	            "POS3_0_Signal"."-1002T1 Oriental_Steuerung".E_DDO_Pos := LREAL_TO_REAL("HMI_COM".HMI_Achse_Steuerung.E_Sollwert_Manuell);
	            "POS3_0_Signal"."-1002T1 Oriental_Steuerung".E_Schrittweite := LREAL_TO_REAL("HMI_COM".HMI_Achse_Steuerung.E_Verfahrweg);
	            "POS3_0_Signal"."-1002T1 Oriental_Steuerung".E_DDO_Vel := LREAL_TO_REAL("HMI_COM".HMI_Achse_Steuerung.E_Geschwindigkeit_manuell_in_Prozent);
	            "POS3_0_Signal"."-1002T1 Oriental_Steuerung".E_DDO_Acc := 100.0;
	            "POS3_0_Signal"."-1002T1 Oriental_Steuerung".E_DDO_Dec := 100.0;
	            "POS3_0_Signal"."-1002T1 Oriental_Steuerung".E_DDO_Crnt := 100;
	            
	            "POS3_0_Signal"."-1002T1 Oriental_Steuerung".E_Schrittweite_pos := "HMI_COM".HMI_Achse_Steuerung.E_Tipp_pos;
	            "POS3_0_Signal"."-1002T1 Oriental_Steuerung".E_Schrittweite_neg := "HMI_COM".HMI_Achse_Steuerung.E_Tipp_neg;
	            "POS3_0_Signal"."-1002T1 Oriental_Steuerung".E_Trig_Manuell := "HMI_COM".HMI_Achse_Steuerung.E_Start_manuell;
	            "POS3_0_Signal"."-1002T1 Oriental_Steuerung"."E_FW-JOG" := "HMI_COM".HMI_Achse_Steuerung.E_jog_pos;
	            "POS3_0_Signal"."-1002T1 Oriental_Steuerung"."E_RV-JOG" := "HMI_COM".HMI_Achse_Steuerung.E_jog_neg;
	        //    "HMI_COM".HMI_Achse_Steuerung.E_Start_manuell := false;
	        END_IF;
	       
	            // Initialisieren der Steuerwerte 
	            #R_TRIG_Init_Achse_2_Positionen(CLK := "HMI_SYS"."Aktueller Bildschirm" = #Manuell_Positionen_1_Achse_2);
	        IF #R_TRIG_Init_Achse_2_Positionen.Q THEN
	                "HMI_COM".HMI_Achse_POS_Überschreiben.Wert_Position_Überschreiben[0] := "POS3_0_Signal"."-1002T1 Oriental_Positionen".Soll_Position[0];
	                "HMI_COM".HMI_Achse_POS_Überschreiben.Wert_Speed_Überschreiben[0] := "POS3_0_Signal"."-1002T1 Oriental_Positionen".Geschwindigkeit[0];
	                
	                "HMI_COM".HMI_Achse_POS_Überschreiben.Wert_Position_Überschreiben[1] := "POS3_0_Signal"."-1002T1 Oriental_Positionen".Soll_Position[1];
	                "HMI_COM".HMI_Achse_POS_Überschreiben.Wert_Speed_Überschreiben[1] := "POS3_0_Signal"."-1002T1 Oriental_Positionen".Geschwindigkeit[1];
	                
	                "HMI_COM".HMI_Achse_POS_Überschreiben.Wert_Position_Überschreiben[2] := "POS3_0_Signal"."-1002T1 Oriental_Positionen".Soll_Position[2];
	                "HMI_COM".HMI_Achse_POS_Überschreiben.Wert_Speed_Überschreiben[2] := "POS3_0_Signal"."-1002T1 Oriental_Positionen".Geschwindigkeit[2];
	                
	                "HMI_COM".HMI_Achse_POS_Überschreiben.Wert_Position_Überschreiben[3] := "POS3_0_Signal"."-1002T1 Oriental_Positionen".Soll_Position[3];
	                "HMI_COM".HMI_Achse_POS_Überschreiben.Wert_Speed_Überschreiben[3] := "POS3_0_Signal"."-1002T1 Oriental_Positionen".Geschwindigkeit[3];
	                
	                "HMI_COM".HMI_Achse_POS_Überschreiben.Wert_Position_Überschreiben[4] := "POS3_0_Signal"."-1002T1 Oriental_Positionen".Soll_Position[4];
	                "HMI_COM".HMI_Achse_POS_Überschreiben.Wert_Speed_Überschreiben[4] := "POS3_0_Signal"."-1002T1 Oriental_Positionen".Geschwindigkeit[4];
	                
	                "HMI_COM".HMI_Achse_POS_Überschreiben.Wert_Position_Überschreiben[5] := "POS3_0_Signal"."-1002T1 Oriental_Positionen".Soll_Position[5];
	                "HMI_COM".HMI_Achse_POS_Überschreiben.Wert_Speed_Überschreiben[5] := "POS3_0_Signal"."-1002T1 Oriental_Positionen".Geschwindigkeit[5];
	        END_IF;
	            
	            
	        IF ("HMI_SYS"."Aktueller Bildschirm" = #Manuell_Positionen_1_Achse_2) THEN
	            
	            "HMI_COM".HMI_Achse_Steuerung.A_StatusWord := "POS3_0_Signal"."-1002T1 Oriental_Steuerung".A_StatusWord;
	            "HMI_COM".HMI_Achse_Steuerung.E_Drehachse := false;
	            "HMI_COM".HMI_Achse_Steuerung.A_Istwert := REAL_TO_LREAL("POS3_0_Signal"."-1002T1 Oriental_Steuerung".A_FBposition);
	            "HMI_COM".HMI_Achse_Steuerung.A_Softw_ES_min := "POS3_0_Signal"."-1002T1 Oriental_Positionen".A_Softw_ES_min_mm;
	            "HMI_COM".HMI_Achse_Steuerung.A_Softw_ES_max := "POS3_0_Signal"."-1002T1 Oriental_Positionen".A_Softw_ES_max_mm;
	            
	            
	            "HMI_COM".HMI_Achse_Position.Soll_Wert_in_mm_Position[0] := "POS3_0_Signal"."-1002T1 Oriental_Positionen".Soll_Position[0];
	            "HMI_COM".HMI_Achse_Position.Soll_Wert_in_mm_Position[1] := "POS3_0_Signal"."-1002T1 Oriental_Positionen".Soll_Position[1];
	            "HMI_COM".HMI_Achse_Position.Soll_Wert_in_mm_Position[2] := "POS3_0_Signal"."-1002T1 Oriental_Positionen".Soll_Position[2];
	            "HMI_COM".HMI_Achse_Position.Soll_Wert_in_mm_Position[3] := "POS3_0_Signal"."-1002T1 Oriental_Positionen".Soll_Position[3];
	            "HMI_COM".HMI_Achse_Position.Soll_Wert_in_mm_Position[4] := "POS3_0_Signal"."-1002T1 Oriental_Positionen".Soll_Position[4];
	            "HMI_COM".HMI_Achse_Position.Soll_Wert_in_mm_Position[5] := "POS3_0_Signal"."-1002T1 Oriental_Positionen".Soll_Position[5];
	            
	            "HMI_COM".HMI_Achse_Position.POS_OK_Position[0] := "POS3_0_Signal"."-1002T1 Oriental_Positionen".POS_OK_Position[0];
	            "HMI_COM".HMI_Achse_Position.POS_OK_Position[1] := "POS3_0_Signal"."-1002T1 Oriental_Positionen".POS_OK_Position[1];
	            "HMI_COM".HMI_Achse_Position.POS_OK_Position[2] := "POS3_0_Signal"."-1002T1 Oriental_Positionen".POS_OK_Position[2];
	            "HMI_COM".HMI_Achse_Position.POS_OK_Position[3] := "POS3_0_Signal"."-1002T1 Oriental_Positionen".POS_OK_Position[3];
	            "HMI_COM".HMI_Achse_Position.POS_OK_Position[4] := "POS3_0_Signal"."-1002T1 Oriental_Positionen".POS_OK_Position[4];
	            "HMI_COM".HMI_Achse_Position.POS_OK_Position[5] := "POS3_0_Signal"."-1002T1 Oriental_Positionen".POS_OK_Position[5];
	            
	            "HMI_COM".HMI_Achse_Position.Soll_Speed_in_Prozent_Position[0] := "POS3_0_Signal"."-1002T1 Oriental_Positionen".Geschwindigkeit[0];
	            "HMI_COM".HMI_Achse_Position.Soll_Speed_in_Prozent_Position[1] := "POS3_0_Signal"."-1002T1 Oriental_Positionen".Geschwindigkeit[1];
	            "HMI_COM".HMI_Achse_Position.Soll_Speed_in_Prozent_Position[2] := "POS3_0_Signal"."-1002T1 Oriental_Positionen".Geschwindigkeit[2];
	            "HMI_COM".HMI_Achse_Position.Soll_Speed_in_Prozent_Position[3] := "POS3_0_Signal"."-1002T1 Oriental_Positionen".Geschwindigkeit[3];
	            "HMI_COM".HMI_Achse_Position.Soll_Speed_in_Prozent_Position[4] := "POS3_0_Signal"."-1002T1 Oriental_Positionen".Geschwindigkeit[4];
	            "HMI_COM".HMI_Achse_Position.Soll_Speed_in_Prozent_Position[5] := "POS3_0_Signal"."-1002T1 Oriental_Positionen".Geschwindigkeit[5];
	            
	            "POS3_0_Signal"."-1002T1 Oriental_Positionen".Start_POS_Position[0] := "HMI_COM".HMI_Achse_Position.Start_POS_Position[0];
	            "POS3_0_Signal"."-1002T1 Oriental_Positionen".Start_POS_Position[1] := "HMI_COM".HMI_Achse_Position.Start_POS_Position[1];
	            "POS3_0_Signal"."-1002T1 Oriental_Positionen".Start_POS_Position[2] := "HMI_COM".HMI_Achse_Position.Start_POS_Position[2];
	            "POS3_0_Signal"."-1002T1 Oriental_Positionen".Start_POS_Position[3] := "HMI_COM".HMI_Achse_Position.Start_POS_Position[3];
	            "POS3_0_Signal"."-1002T1 Oriental_Positionen".Start_POS_Position[4] := "HMI_COM".HMI_Achse_Position.Start_POS_Position[4];
	            "POS3_0_Signal"."-1002T1 Oriental_Positionen".Start_POS_Position[5] := "HMI_COM".HMI_Achse_Position.Start_POS_Position[5];
	        
	            
	            IF "HMI_COM".HMI_Achse_POS_Überschreiben.Trig_Position_Überschreiben[0] THEN
	                "POS3_0_Signal"."-1002T1 Oriental_Positionen".Soll_Position[0] := "HMI_COM".HMI_Achse_POS_Überschreiben.Wert_Position_Überschreiben[0];
	                "POS3_0_Signal"."-1002T1 Oriental_Positionen".Geschwindigkeit[0] := "HMI_COM".HMI_Achse_POS_Überschreiben.Wert_Speed_Überschreiben[0];
	            END_IF;
	            
	            IF "HMI_COM".HMI_Achse_POS_Überschreiben.Trig_Position_Überschreiben[1] THEN
	                "POS3_0_Signal"."-1002T1 Oriental_Positionen".Soll_Position[1] := "HMI_COM".HMI_Achse_POS_Überschreiben.Wert_Position_Überschreiben[1];
	                "POS3_0_Signal"."-1002T1 Oriental_Positionen".Geschwindigkeit[1] := "HMI_COM".HMI_Achse_POS_Überschreiben.Wert_Speed_Überschreiben[1];
	            END_IF;
	            
	            IF "HMI_COM".HMI_Achse_POS_Überschreiben.Trig_Position_Überschreiben[2] THEN
	                "POS3_0_Signal"."-1002T1 Oriental_Positionen".Soll_Position[2] := "HMI_COM".HMI_Achse_POS_Überschreiben.Wert_Position_Überschreiben[2];
	                "POS3_0_Signal"."-1002T1 Oriental_Positionen".Geschwindigkeit[2] := "HMI_COM".HMI_Achse_POS_Überschreiben.Wert_Speed_Überschreiben[2];
	            END_IF;
	            
	            IF "HMI_COM".HMI_Achse_POS_Überschreiben.Trig_Position_Überschreiben[3] THEN
	                "POS3_0_Signal"."-1002T1 Oriental_Positionen".Soll_Position[3] := "HMI_COM".HMI_Achse_POS_Überschreiben.Wert_Position_Überschreiben[3];
	                "POS3_0_Signal"."-1002T1 Oriental_Positionen".Geschwindigkeit[3] := "HMI_COM".HMI_Achse_POS_Überschreiben.Wert_Speed_Überschreiben[3];
	            END_IF;
	            
	            IF "HMI_COM".HMI_Achse_POS_Überschreiben.Trig_Position_Überschreiben[4] THEN
	                "POS3_0_Signal"."-1002T1 Oriental_Positionen".Soll_Position[4] := "HMI_COM".HMI_Achse_POS_Überschreiben.Wert_Position_Überschreiben[4];
	                "POS3_0_Signal"."-1002T1 Oriental_Positionen".Geschwindigkeit[4] := "HMI_COM".HMI_Achse_POS_Überschreiben.Wert_Speed_Überschreiben[4];
	            END_IF;
	            
	            IF "HMI_COM".HMI_Achse_POS_Überschreiben.Trig_Position_Überschreiben[5] THEN
	                "POS3_0_Signal"."-1002T1 Oriental_Positionen".Soll_Position[5] := "HMI_COM".HMI_Achse_POS_Überschreiben.Wert_Position_Überschreiben[5];
	                "POS3_0_Signal"."-1002T1 Oriental_Positionen".Geschwindigkeit[5] := "HMI_COM".HMI_Achse_POS_Überschreiben.Wert_Speed_Überschreiben[5];
	            END_IF;
	            
	        END_IF;
	        
	        IF ("HMI_SYS"."Aktueller Bildschirm" = #"Manuell_P-Preset_1_Achse_2") THEN
	            "HMI_COM".HMI_Achse_Steuerung.A_StatusWord := "POS3_0_Signal"."-1002T1 Oriental_Steuerung".A_StatusWord;
	            "HMI_COM".HMI_Achse_Steuerung.E_Drehachse := true;
	            "HMI_COM".HMI_Achse_Steuerung.A_Istwert := REAL_TO_LREAL("POS3_0_Signal"."-1002T1 Oriental_Steuerung".A_FBposition);
	        END_IF;
	        
	        
	    END_REGION
	    
	    
	    
	    
	END_REGION
	
	
	
	
	
	
END_FUNCTION_BLOCK

FUNCTION_BLOCK "Taktzeitermittlung_Start_Stop_V1_0"
TITLE = Taktzeitermittlung Start Stop
{ S7_Optimized_Access := 'TRUE' }
AUTHOR : FA
VERSION : 1.0
//Ausgabe der Zeit zwischen 1 und 0 Signal am Starttrigger 27.03.2024 FA
   VAR_INPUT 
      E_Starttrigger : Bool;
   END_VAR

   VAR_OUTPUT 
      A_letzteZykluszeit : Time;
   END_VAR
   VAR_OUTPUT DB_SPECIFIC
      A_letze10Zyklen : Array[0..10] of Time := [T#1MS, T#765MS, T#759MS, T#762MS, T#758MS, T#763MS, T#768MS, T#763MS, T#766MS, T#757MS, T#766MS];
   END_VAR

   VAR 
      Flanke_Start {InstructionName := 'R_TRIG'; LibVersion := '1.0'} : R_TRIG;
      Flanke_Stop {InstructionName := 'F_TRIG'; LibVersion := '1.0'} : F_TRIG;
      Startzeit { S7_SetPoint := 'True'} : LDT;
      Stopzeit : LDT;
      Read_Time : Int;
      Taktzeit : Time;
      Zykluszeit_temp : Time;
      "10_Zyklen" : Array[0..10] of Time;
   END_VAR

   VAR_TEMP 
      i : Int;
   END_VAR


BEGIN
	(*
	Zeit zwischen Positiver und negativer Flanke am Triggereingang wird ermittelt und am Ausgang letzte Zykluszeit ausgegeben
	zusätzlichwerden die letzten 10 Zykluszeiten am Ausgangangsarray ausgegeben *)
	
	#Flanke_Start(CLK := #E_Starttrigger);
	    #Flanke_Stop(CLK := #E_Starttrigger);
	    
	    IF #Flanke_Start.Q THEN
	     
	        #Read_Time := RD_SYS_T(#Startzeit);
	    
	       
	    END_IF;
	    
	    
	    IF #Flanke_Stop.Q THEN
	        #Read_Time := RD_SYS_T(#Stopzeit);
	        
	        #Taktzeit := LTIME_TO_TIME(LDT_TO_LTIME(T_SUB(IN1 := #Stopzeit, IN2 :=#Startzeit)));
	        #"10_Zyklen"[0] := #Taktzeit;
	        FOR #i := 10 TO 1 BY - 1 DO
	            #"10_Zyklen"[#i] := #"10_Zyklen"[#i - 1]
	            ;
	        END_FOR;
	        
	        #A_letzteZykluszeit := #"10_Zyklen"[1];
	        #A_letze10Zyklen := #"10_Zyklen";
	        
	        #Zykluszeit_temp := t#0s;
	        #Stopzeit := #Startzeit;
	    END_IF;
	    
END_FUNCTION_BLOCK

FUNCTION "POS3_0_Teileauswertung" : Void   // FC60, STL
TITLE = Teileauswertung
{ S7_Optimized_Access := 'FALSE' }
   VAR_TEMP
      RetVal : Int;
   END_VAR
BEGIN
END_FUNCTION

FUNCTION_BLOCK "POS3_0_Messtechnik"
{ S7_Optimized_Access := 'TRUE' }
VERSION : 0.1

BEGIN
	
	
	 
	REGION -1012B1 Kraftsensor
	    
	    "POS3_0_Signal"."-1012B1 Kraftsensor" := DWORD_TO_REAL("IN-POS3_0-1012B1 Kraftsensor");
	END_REGION
	
	
	REGION -940RN1 Regelventil Ausgleichszylinder
	    // Vorgabe der maximalen Abweichung; evtl. aus Programmvorgabe !!!
	    "POS3_0_Signal"."-POS3_0_Regelventil_Ausgleichszylinder_Maximale_Abweichung" := 100;
	    
	    "IO-OUT-POS3_0_Regelventil_Ausgleichszylinder_Sollwert"   := "POS3_0_Signal"."-POS3_0_Regelventil_Ausgleichszylinder_Sollwert";
	    "POS3_0_Signal"."-POS3_0_Regelventil_Ausgleichszylinder_Istwert" := "IO-IN-POS3_0_Regelventil_Ausgleichszylinder_Istwert";
	    
	    REGION Maximale Regelabweichung       
	        "POS3_0_Signal"."-POS3_0_Regelventil_Ausgleichszylinder_Abweichung_OK" :=
	        ABS(
	            "POS3_0_Signal"."-POS3_0_Regelventil_Ausgleichszylinder_Istwert" - "POS3_0_Signal"."-POS3_0_Regelventil_Ausgleichszylinder_Sollwert")
	        <= "POS3_0_Signal"."-POS3_0_Regelventil_Ausgleichszylinder_Maximale_Abweichung";
	    END_REGION
	    
	END_REGION
	
	
	
	REGION -940RN2 Regelventil Überlastzylinder
	    // Vorgabe der maximalen Abweichung; evtl. aus Programmvorgabe !!!
	    "POS3_0_Signal"."-POS3_0_Regelventil_Überlastzylinder_Maximale_Abweichung" := 100;
	    
	    "IO-OUT-POS3_0_Regelventil_Überlastzylinder_Sollwert" := "POS3_0_Signal"."-POS3_0_Regelventil_Überlastzylinder_Sollwert";
	    "POS3_0_Signal"."-POS3_0_Regelventil_Überlastzylinder_Istwert" := "IO-IN-POS3_0_Regelventil_Überlastzylinder_Istwert";
	    
	    REGION Maximale Regelabweichung
	        "POS3_0_Signal"."-POS3_0_Regelventil_Überlastzylinder_Abweichung_OK" :=
	        ABS(
	            "POS3_0_Signal"."-POS3_0_Regelventil_Überlastzylinder_Istwert" - "POS3_0_Signal"."-POS3_0_Regelventil_Überlastzylinder_Sollwert")
	        <= "POS3_0_Signal"."-POS3_0_Regelventil_Überlastzylinder_Maximale_Abweichung";
	    END_REGION
	    
	END_REGION
	
	
	REGION Wegmessung Ausgleichszylinder
	    // Rohwert 
	    "POS3_0_Signal"."-POS3.0_Wegmessung_Ausgleichszylinder_Istwert_Rohwert" := "IO-IN-POS3_0_Wegmessung_Ausgleichszylinder_Istwert";
	    
	    // Taster Nullen
	    IF "POS3_0_Signal"."-POS3.0_Wegmessung_Ausgleichszylinder_Taster_Nullen" THEN
	        "POS3_0_Signal"."-POS3.0_Wegmessung_Ausgleichszylinder_Nullpunkt_Rohwert" := "POS3_0_Signal"."-POS3.0_Wegmessung_Ausgleichszylinder_Istwert_Rohwert";
	        "POS3_0_Signal"."-POS3.0_Wegmessung_Ausgleichszylinder_Taster_Nullen" := false;
	    END_IF;
	    
	    // Normierung
	    "POS3_0_Signal"."-POS3.0_Wegmessung_Ausgleichszylinder_Istwert_in_mm" :=
	    (INT_TO_REAL("POS3_0_Signal"."-POS3.0_Wegmessung_Ausgleichszylinder_Istwert_Rohwert" - "POS3_0_Signal"."-POS3.0_Wegmessung_Ausgleichszylinder_Nullpunkt_Rohwert"))
	    * 38.5 / 12624.0;
	    
	    
	    
	    REGION Maximale Abweichung GS
	        "POS3_0_Signal"."-POS3.0_Wegmessung_Ausgleichszylinder_Position_GS_Abweichung_OK" :=
	        ABS(
	            "POS3_0_Signal"."-POS3.0_Wegmessung_Ausgleichszylinder_Istwert_in_mm" - "Verwaltung_Teiledaten"."Wegmessung_Ausgleichszylinder Position GS")
	        <= "Verwaltung_Teiledaten"."Wegmessung_Ausgleichszylinder maximale Abweichung GS";
	    END_REGION
	    
	    
	    
	    REGION Maximale Abweichung AS1
	        "POS3_0_Signal"."-POS3.0_Wegmessung_Ausgleichszylinder_Position_AS1_Abweichung_OK" :=
	        ABS(
	            "POS3_0_Signal"."-POS3.0_Wegmessung_Ausgleichszylinder_Istwert_in_mm" - "Verwaltung_Teiledaten"."Wegmessung_Ausgleichszylinder Position AS1")
	        <= "Verwaltung_Teiledaten"."Wegmessung_Ausgleichszylinder maximale Abweichung AS1";
	    END_REGION
	    
	    
	END_REGION
	
	
END_FUNCTION_BLOCK

FUNCTION_BLOCK "POS3_0_SK_Ablauf"   // FB26, GRAPH
// stored: GraphVersion 6.0, InitialValuesAcquisition false, LanguageInNetworks FBD, SetENOAutomatically false
   // inherited from GRAPH_BASE
   VAR_INPUT
      OFF_SQ { ExternalWritable := 'False'} : Bool := false;   // Kette ausschalten
      INIT_SQ { ExternalWritable := 'False'} : Bool := false;   // Kette in Initialzustand versetzen
      ACK_EF { ExternalWritable := 'False'} : Bool := false;   // Alle Fehler und Störungen quittieren
      REG_EF { ExternalWritable := 'False'} : Bool := false;   // Alle Fehler und Störungen registrieren
      ACK_S { ExternalWritable := 'False'} : Bool := false;   // Schritt quittieren, der an Parameter S_NO anliegt
      REG_S { ExternalWritable := 'False'} : Bool := false;   // Schritt registrieren, der an Parameter S_NO anliegt
      HALT_SQ { ExternalWritable := 'False'} : Bool := false;   // Kette sofort anhalten
      HALT_TM { ExternalWritable := 'False'} : Bool := false;   // Zeiten sofort anhalten
      ZERO_OP { ExternalWritable := 'False'} : Bool := false;   // Alle mit N, L, D zugewiesenen Operanden auf 0 setzen
      EN_IL { ExternalWritable := 'False'} : Bool := false;   // Interlockbearbeitung aktivieren
      EN_SV { ExternalWritable := 'False'} : Bool := false;   // Supervisionsbearbeitung aktivieren
      EN_ACKREQ { ExternalWritable := 'False'} : Bool := false;   // Quittierpflicht aktivieren
      EN_SSKIP { ExternalWritable := 'False'} : Bool := false;   // "Schritte überspringen" aktivieren
      DISP_SACT { ExternalWritable := 'False'} : Bool := false;   // Nur aktive Schritte anzeigen
      DISP_SEF { ExternalWritable := 'False'} : Bool := false;   // Nur fehlerhafte und gestörte Schritte anzeigen
      DISP_SALL { ExternalWritable := 'False'} : Bool := false;   // Alle Schritte anzeigen
      S_PREV { ExternalWritable := 'False'} : Bool := false;   // Vorherigen Schritt am Parameter S_NO ausgeben
      S_NEXT { ExternalWritable := 'False'} : Bool := false;   // Nächsten Schritt am Parameter S_NO anzeigen
      SW_AUTO { ExternalWritable := 'False'} : Bool := false;   // Automatischer Betrieb
      SW_TAP { ExternalWritable := 'False'} : Bool := false;   // Halbautomatisch/Weiterschalten mit Transition
      SW_TOP { ExternalWritable := 'False'} : Bool := false;   // Halbautomatisch/Ignoriere Transition
      SW_MAN { ExternalWritable := 'False'} : Bool := false;   // Handbetrieb
      S_SEL { ExternalWritable := 'False'} : Int := 0;   // Schritt auswählen, der an S_NO ausgegeben werden soll
      S_SELOK { ExternalWritable := 'False'} : Bool := false;   // Wert aus S_SEL nach S_NO übernehmen
      S_ON { ExternalWritable := 'False'} : Bool := false;   // Schritt aktivieren, der an Parameter S_NO anliegt
      S_OFF { ExternalWritable := 'False'} : Bool := false;   // Schritt deaktivieren, der an Parameter S_NO anliegt
      T_PREV { ExternalWritable := 'False'} : Bool := false;   // Vorherige Transition an Parameter T_NO anzeigen
      T_NEXT { ExternalWritable := 'False'} : Bool := false;   // Nächste Transition an Parameter T_NO anzeigen
      T_PUSH { ExternalWritable := 'False'} : Bool := false;   // Schaltfreigabe für Transition im halbautomatischen Betrieb
      EN_LMODE { ExternalWritable := 'False'} : Bool := false;   // Lernmodus aktivieren
   END_VAR
   VAR_OUTPUT
      S_NO { ExternalWritable := 'False'} : Int := 0;   // Schrittnummer
      S_MORE { ExternalWritable := 'False'} : Bool := false;   // Weitere Schritte sind vorhanden und können in S_NO angezeigt werden.
      S_ACTIVE { ExternalWritable := 'False'} : Bool := false;   // Schritt, der an Parameter S_NO angezeigt wird, ist aktiv
      S_TIME { ExternalWritable := 'False'} : Time := T#0ms;   // Schrittaktivierungszeit
      S_TIMEOK { ExternalWritable := 'False'} : Time := T#0ms;   // Schrittaktivierungszeit fehlerfrei
      S_CRITLOC { ExternalWritable := 'False'} : DWord := 16#0;   // Interlock-Kriterienbits
      S_CRITLOCERR { ExternalWritable := 'False'} : DWord := 16#0;   // Interlock-Kriterienbits bei Ereignis L1
      S_STATE { ExternalWritable := 'False'} : Word := 16#0;   // Schrittzustandsbits
      T_NO { ExternalWritable := 'False'} : Int := 0;   // Transitionsnummer
      T_MORE { ExternalWritable := 'False'} : Bool := false;   // Weitere gültige Transitionen zur Anzeige verfügbar
      T_CRIT { ExternalWritable := 'False'} : DWord := 16#0;   // Transitions-Kriterienbits
      T_CRITOLD { ExternalWritable := 'False'} : DWord := 16#0;   // Transitions-Kriterienbits des letzten Zyklus
      T_CRITFLT { ExternalWritable := 'False'} : DWord := 16#0;   // Transitions-Kriterienbits bei Ereignis V1
      ERROR { ExternalWritable := 'False'} : Bool := false;   // Sammelfehler Interlock
      FAULT { ExternalWritable := 'False'} : Bool := false;   // Sammelfehler Supervision
      ERR_FLT { ExternalWritable := 'False'} : Bool := false;   // Sammelfehler Interlock oder Supervision
      SQ_ISOFF { ExternalWritable := 'False'} : Bool := false;   // Kette ausgeschaltet (kein Schritt aktiv)
      SQ_HALTED { ExternalWritable := 'False'} : Bool := false;   // Kette angehalten
      TM_HALTED { ExternalWritable := 'False'} : Bool := false;   // Zeiten angehalten
      OP_ZEROED { ExternalWritable := 'False'} : Bool := false;   // Alle mit N, L oder D zugewiesenen Operanden auf 0 gesetzt
      IL_ENABLED { ExternalWritable := 'False'} : Bool := false;   // Interlockbearbeitung aktiv
      SV_ENABLED { ExternalWritable := 'False'} : Bool := false;   // Supervisionsbearbeitung aktiviert
      ACKREQ_ENABLED { ExternalWritable := 'False'} : Bool := false;   // Quittierpflicht aktiviert
      SSKIP_ENABLED { ExternalWritable := 'False'} : Bool := false;   // Schritte überspringen aktiviert
      SACT_DISP { ExternalWritable := 'False'} : Bool := false;   // Nur aktive Schritte anzeigen
      SEF_DISP { ExternalWritable := 'False'} : Bool := false;   // Nur fehlerhafte oder gestörte Schritte anzeigen
      SALL_DISP { ExternalWritable := 'False'} : Bool := false;   // Alle Schritte anzeigen
      AUTO_ON { ExternalWritable := 'False'} : Bool := false;   // Automatischer Betrieb eingeschaltet
      TAP_ON { ExternalWritable := 'False'} : Bool := false;   // Halbautomatischer Betrieb/Schritt mit Transition eingeschaltet
      TOP_ON { ExternalWritable := 'False'} : Bool := false;   // Halbautomatischer Betrieb/Ignoriere Transition eingeschaltet
      MAN_ON { ExternalWritable := 'False'} : Bool := false;   // Handbetrieb eingeschaltet
      LMODE_ENABLED { ExternalWritable := 'False'} : Bool := false;   // Lernmodus aktiv
   END_VAR
BEGIN
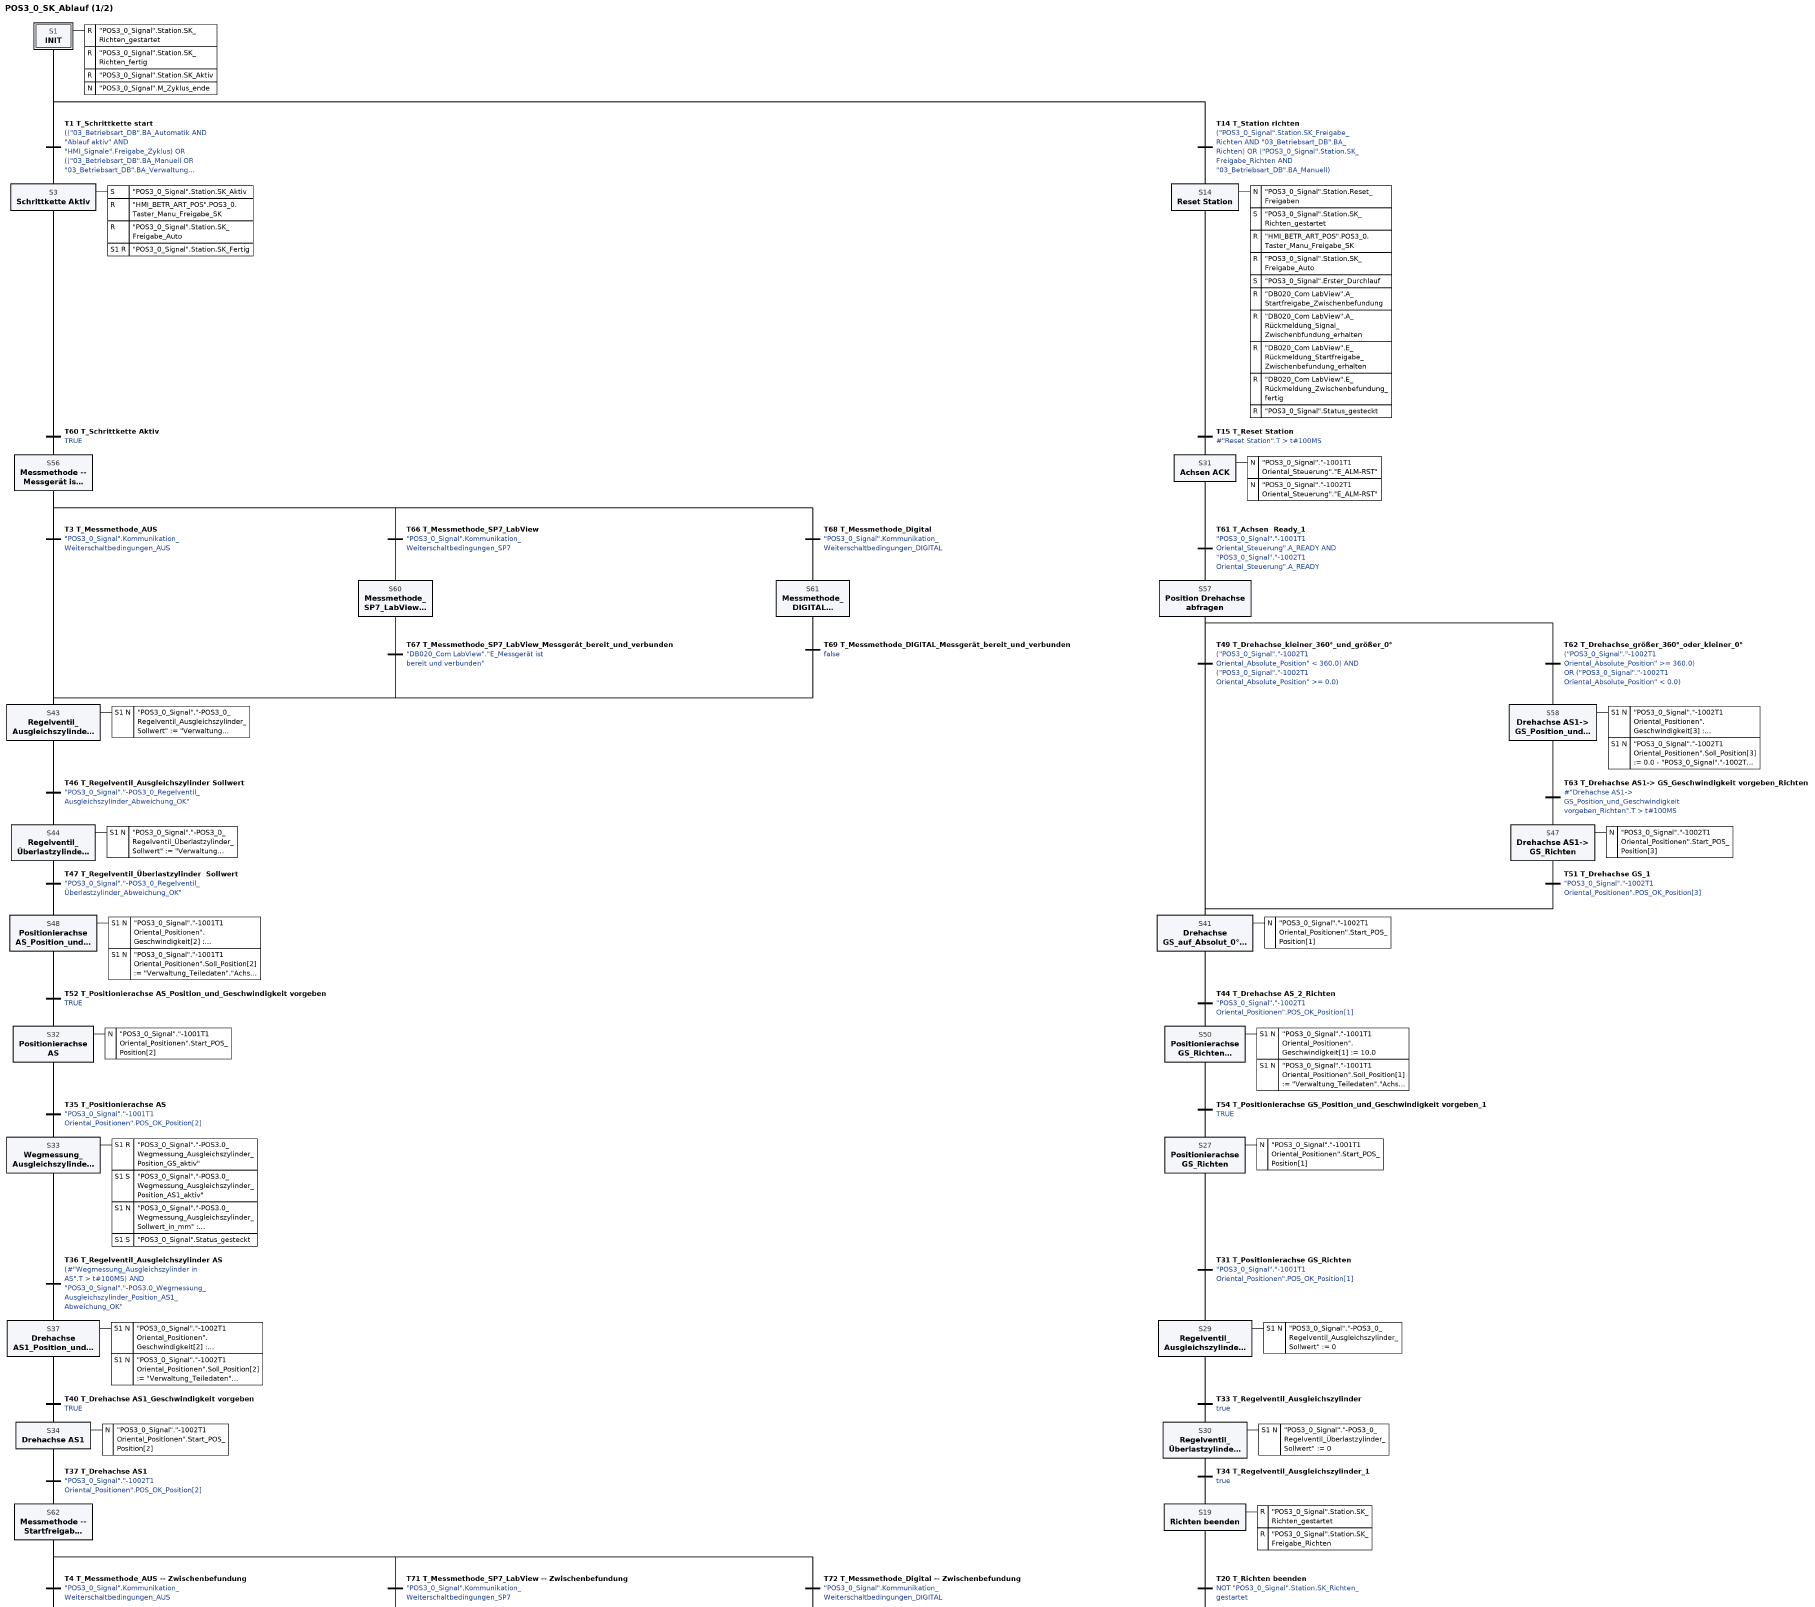
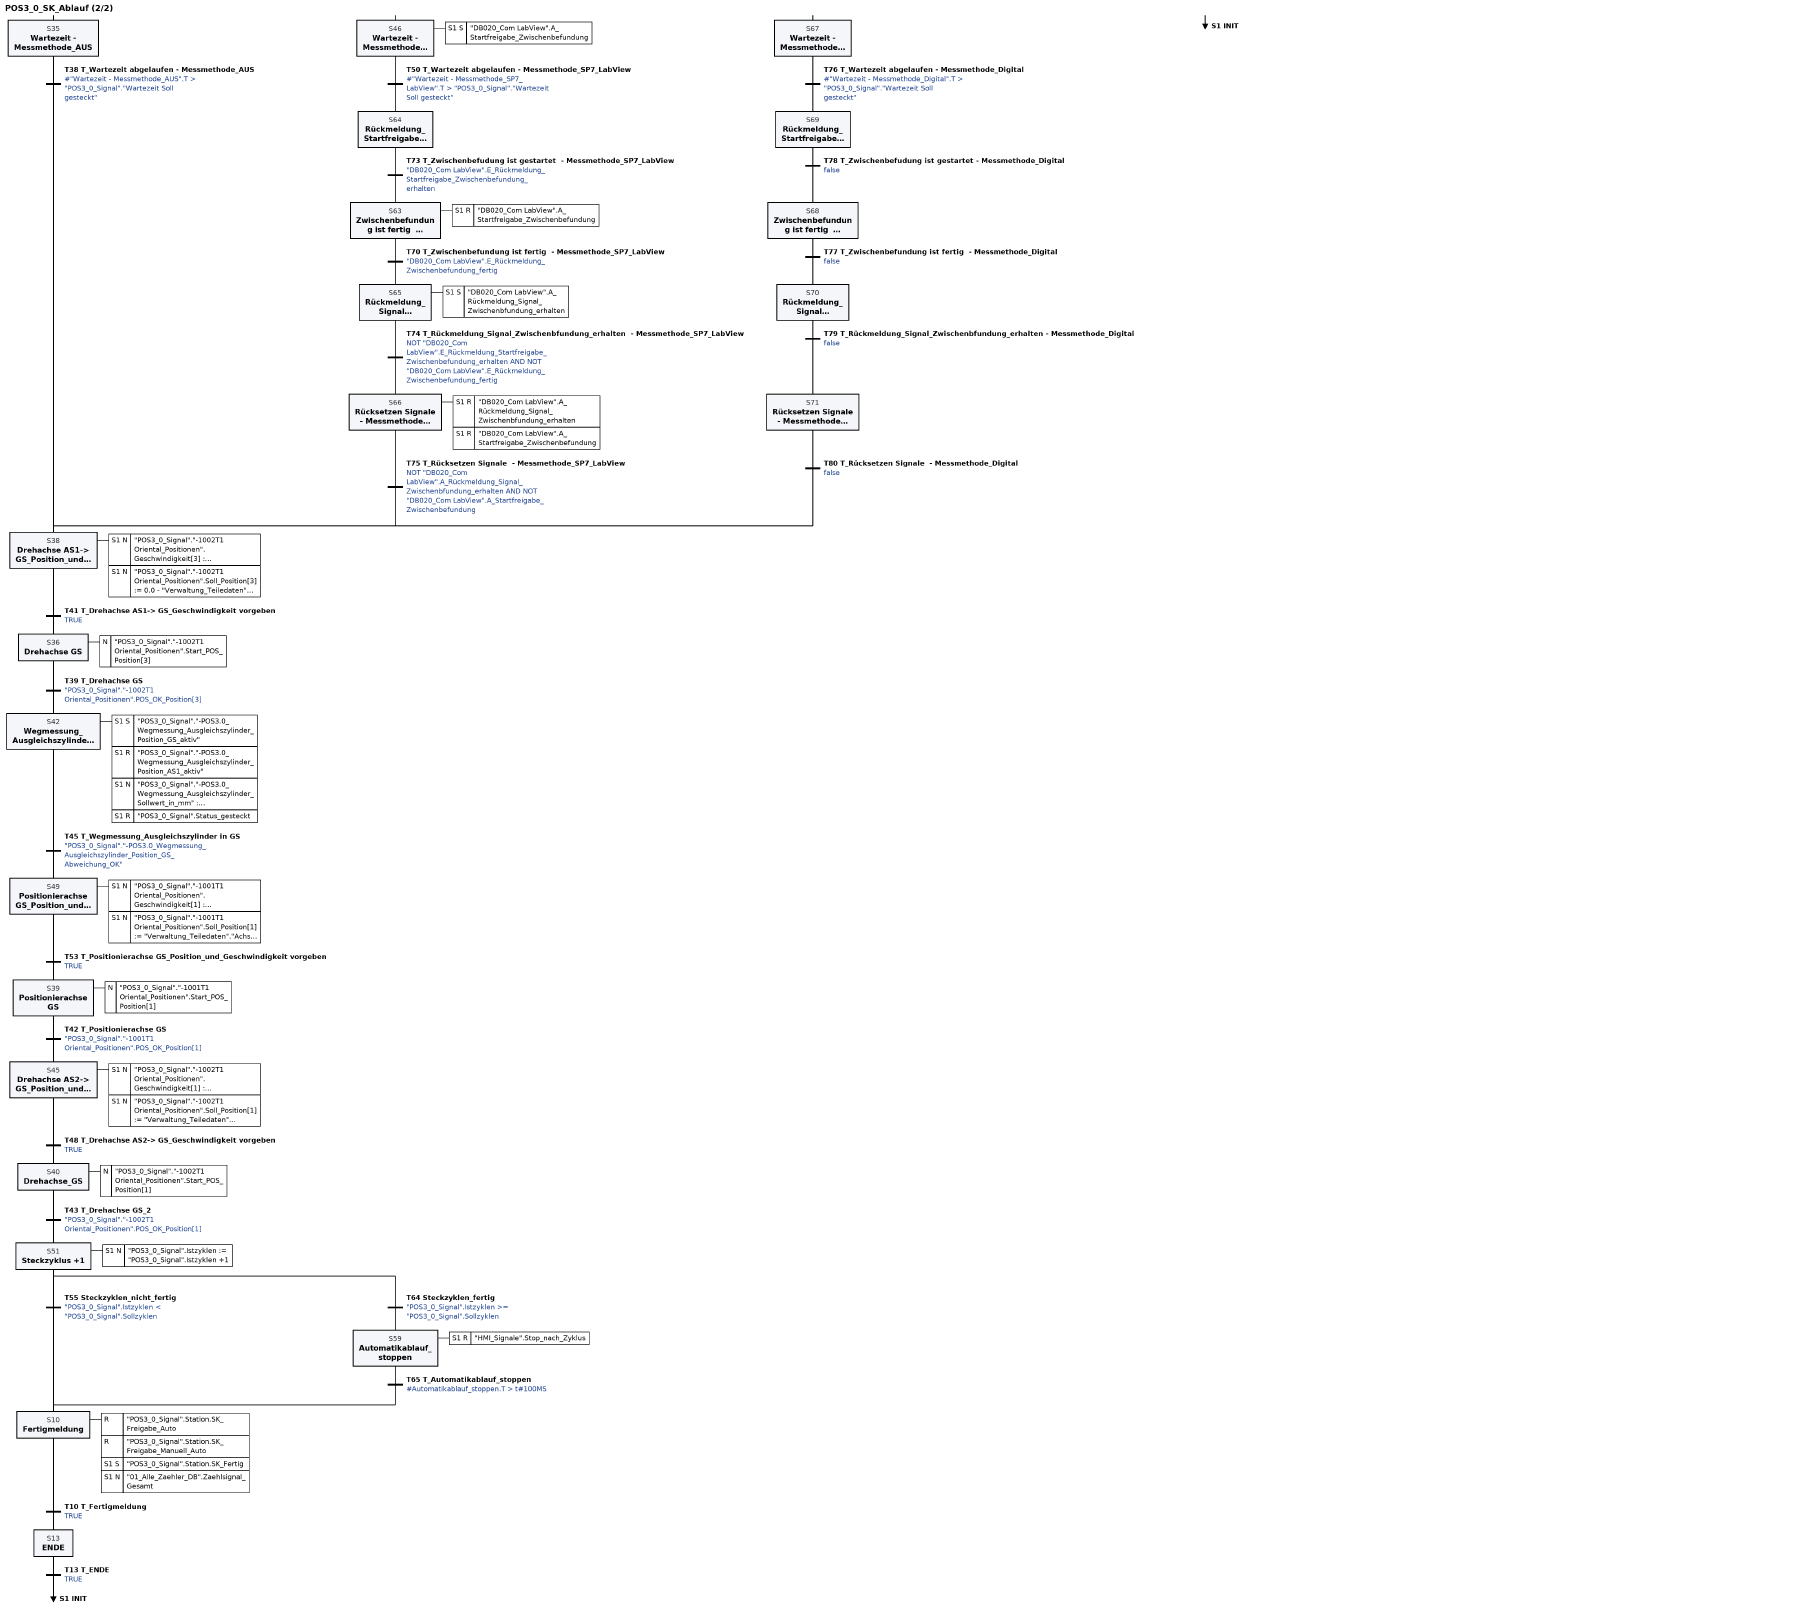
   // sequencer 1
   INITIAL_STEP INIT:   // S1, max time T#10S, warning time T#7S
              R    "POS3_0_Signal".Station.SK_Richten_gestartet
              R    "POS3_0_Signal".Station.SK_Richten_fertig
              R    "POS3_0_Signal".Station.SK_Aktiv
              N    "POS3_0_Signal".M_Zyklus_ende
   END_STEP
   TRANSITION "T_Schrittkette start" FROM INIT TO "Schrittkette Aktiv"   // T1
      := (("03_Betriebsart_DB".BA_Automatik AND "Ablauf aktiv" AND "HMI_Signale".Freigabe_Zyklus) OR (("03_Betriebsart_DB".BA_Manuell OR "03_Betriebsart_DB".BA_Verwaltung) AND "HMI_BETR_ART_POS".POS3_0.Taster_Manu_Freigabe_SK)) AND "Global_Signal"."M_Grundstellung_POS3.0";
   END_TRANSITION
   TRANSITION "T_Station richten" FROM INIT TO "Reset Station"   // T14
      := ("POS3_0_Signal".Station.SK_Freigabe_Richten AND "03_Betriebsart_DB".BA_Richten) OR ("POS3_0_Signal".Station.SK_Freigabe_Richten AND "03_Betriebsart_DB".BA_Manuell);
   END_TRANSITION
   STEP "Schrittkette Aktiv":   // S3, max time T#10S, warning time T#7S
      supervision V := #"Schrittkette Aktiv".U > #"Schrittkette Aktiv".T_MAX;
              S    "POS3_0_Signal".Station.SK_Aktiv
              R    "HMI_BETR_ART_POS".POS3_0.Taster_Manu_Freigabe_SK
              R    "POS3_0_Signal".Station.SK_Freigabe_Auto
          S1  R    "POS3_0_Signal".Station.SK_Fertig
   END_STEP
   TRANSITION "T_Schrittkette Aktiv" FROM "Schrittkette Aktiv" TO "Messmethode -- Messgerät ist bereit oder nicht verbunden"   // T60
      := TRUE;
   END_TRANSITION
   STEP "Drehachse GS":   // S36, max time T#10S, warning time T#7S
      supervision V := #"Drehachse GS".U > #"Drehachse GS".T_MAX;
              N    "POS3_0_Signal"."-1002T1 Oriental_Positionen".Start_POS_Position[3]
   END_STEP
   TRANSITION "T_Drehachse GS" FROM "Drehachse GS" TO "Wegmessung_Ausgleichszylinder in GS"   // T39
      := "POS3_0_Signal"."-1002T1 Oriental_Positionen".POS_OK_Position[3];
   END_TRANSITION
   STEP Fertigmeldung:   // S10, max time T#10S, warning time T#7S
      supervision V := #Fertigmeldung.U > #Fertigmeldung.T_MAX;
              R    "POS3_0_Signal".Station.SK_Freigabe_Auto
              R    "POS3_0_Signal".Station.SK_Freigabe_Manuell_Auto
          S1  S    "POS3_0_Signal".Station.SK_Fertig
          S1  N    "01_Alle_Zaehler_DB".Zaehlsignal_Gesamt
   END_STEP
   TRANSITION T_Fertigmeldung FROM Fertigmeldung TO ENDE   // T10
      := TRUE;
   END_TRANSITION
   STEP ENDE:   // S13, max time T#10S, warning time T#7S
   END_STEP
   TRANSITION T_ENDE FROM ENDE TO INIT   // T13, jump
      := TRUE;
   END_TRANSITION
   STEP "Reset Station":   // S14, max time T#10S, warning time T#7S
              N    "POS3_0_Signal".Station.Reset_Freigaben
              S    "POS3_0_Signal".Station.SK_Richten_gestartet
              R    "HMI_BETR_ART_POS".POS3_0.Taster_Manu_Freigabe_SK
              R    "POS3_0_Signal".Station.SK_Freigabe_Auto
              S    "POS3_0_Signal".Erster_Durchlauf
              R    "DB020_Com LabView".A_Startfreigabe_Zwischenbefundung
              R    "DB020_Com LabView".A_Rückmeldung_Signal_Zwischenbfundung_erhalten
              R    "DB020_Com LabView".E_Rückmeldung_Startfreigabe_Zwischenbefundung_erhalten
              R    "DB020_Com LabView".E_Rückmeldung_Zwischenbefundung_fertig
              R    "POS3_0_Signal".Status_gesteckt
   END_STEP
   TRANSITION "T_Reset Station" FROM "Reset Station" TO "Achsen ACK"   // T15
      := #"Reset Station".T > t#100MS;
   END_TRANSITION
   STEP "Richten beenden":   // S19, max time T#10S, warning time T#7S
              R    "POS3_0_Signal".Station.SK_Richten_gestartet
              R    "POS3_0_Signal".Station.SK_Freigabe_Richten
   END_STEP
   TRANSITION "T_Richten beenden" FROM "Richten beenden" TO INIT   // T20, jump
      := NOT "POS3_0_Signal".Station.SK_Richten_gestartet;
   END_TRANSITION
   STEP "Wartezeit - Messmethode_AUS":   // S35, max time T#10S, warning time T#7S
   END_STEP
   TRANSITION "T_Wartezeit abgelaufen - Messmethode_AUS" FROM "Wartezeit - Messmethode_AUS" TO "Drehachse AS1-> GS_Position_und_Geschwindigkeit vorgeben"   // T38
      := #"Wartezeit - Messmethode_AUS".T > "POS3_0_Signal"."Wartezeit Soll gesteckt";
   END_TRANSITION
   STEP "Positionierachse GS_Richten":   // S27, max time T#10S, warning time T#7S
      supervision V := #"Positionierachse GS_Richten".U > #"Positionierachse GS_Richten".T_MAX;
              N    "POS3_0_Signal"."-1001T1 Oriental_Positionen".Start_POS_Position[1]
   END_STEP
   TRANSITION "T_Positionierachse GS_Richten" FROM "Positionierachse GS_Richten" TO "Regelventil_Ausgleichszylinder auf 0 mbar"   // T31
      := "POS3_0_Signal"."-1001T1 Oriental_Positionen".POS_OK_Position[1];
   END_TRANSITION
   STEP "Achsen ACK":   // S31, max time T#10S, warning time T#7S
              N    "POS3_0_Signal"."-1001T1 Oriental_Steuerung"."E_ALM-RST"
              N    "POS3_0_Signal"."-1002T1 Oriental_Steuerung"."E_ALM-RST"
   END_STEP
   TRANSITION "T_Achsen  Ready_1" FROM "Achsen ACK" TO "Position Drehachse abfragen"   // T61
      := "POS3_0_Signal"."-1001T1 Oriental_Steuerung".A_READY AND "POS3_0_Signal"."-1002T1 Oriental_Steuerung".A_READY;
   END_TRANSITION
   STEP "Regelventil_Ausgleichszylinder auf 0 mbar":   // S29, max time T#10S, warning time T#7S
          S1  N    "POS3_0_Signal"."-POS3_0_Regelventil_Ausgleichszylinder_Sollwert" := 0
   END_STEP
   TRANSITION T_Regelventil_Ausgleichszylinder FROM "Regelventil_Ausgleichszylinder auf 0 mbar" TO "Regelventil_Überlastzylinder auf 0 mbar"   // T33
      := true;
   END_TRANSITION
   STEP "Regelventil_Überlastzylinder auf 0 mbar":   // S30, max time T#10S, warning time T#7S
          S1  N    "POS3_0_Signal"."-POS3_0_Regelventil_Überlastzylinder_Sollwert" := 0
   END_STEP
   TRANSITION T_Regelventil_Ausgleichszylinder_1 FROM "Regelventil_Überlastzylinder auf 0 mbar" TO "Richten beenden"   // T34
      := true;
   END_TRANSITION
   STEP "Positionierachse AS":   // S32, max time T#10S, warning time T#7S
      supervision V := #"Positionierachse AS".U > t#300s;
              N    "POS3_0_Signal"."-1001T1 Oriental_Positionen".Start_POS_Position[2]
   END_STEP
   TRANSITION "T_Positionierachse AS" FROM "Positionierachse AS" TO "Wegmessung_Ausgleichszylinder in AS"   // T35
      := "POS3_0_Signal"."-1001T1 Oriental_Positionen".POS_OK_Position[2];
   END_TRANSITION
   STEP "Wegmessung_Ausgleichszylinder in AS":   // S33, max time T#10S, warning time T#7S
      supervision V := #"Wegmessung_Ausgleichszylinder in AS".U > #"Wegmessung_Ausgleichszylinder in AS".T_MAX;
          S1  R    "POS3_0_Signal"."-POS3.0_Wegmessung_Ausgleichszylinder_Position_GS_aktiv"
          S1  S    "POS3_0_Signal"."-POS3.0_Wegmessung_Ausgleichszylinder_Position_AS1_aktiv"
          S1  N    "POS3_0_Signal"."-POS3.0_Wegmessung_Ausgleichszylinder_Sollwert_in_mm" := "Verwaltung_Teiledaten"."Wegmessung_Ausgleichszylinder Position AS1"
          S1  S    "POS3_0_Signal".Status_gesteckt
   END_STEP
   TRANSITION "T_Regelventil_Ausgleichszylinder AS" FROM "Wegmessung_Ausgleichszylinder in AS" TO "Drehachse AS1_Position_und_Geschwindigkeit vorgeben"   // T36
      := (#"Wegmessung_Ausgleichszylinder in AS".T > t#100MS) AND "POS3_0_Signal"."-POS3.0_Wegmessung_Ausgleichszylinder_Position_AS1_Abweichung_OK";
   END_TRANSITION
   STEP "Drehachse AS1":   // S34, max time T#10S, warning time T#7S
      supervision V := #"Drehachse AS1".U > #"Drehachse AS1".T_MAX;
              N    "POS3_0_Signal"."-1002T1 Oriental_Positionen".Start_POS_Position[2]
   END_STEP
   TRANSITION "T_Drehachse AS1" FROM "Drehachse AS1" TO "Messmethode -- Startfreigabe Zwischenbefundung"   // T37
      := "POS3_0_Signal"."-1002T1 Oriental_Positionen".POS_OK_Position[2];
   END_TRANSITION
   STEP "Positionierachse GS":   // S39, max time T#10S, warning time T#7S
      supervision V := #"Positionierachse GS".U > t#300s;
              N    "POS3_0_Signal"."-1001T1 Oriental_Positionen".Start_POS_Position[1]
   END_STEP
   TRANSITION "T_Positionierachse GS" FROM "Positionierachse GS" TO "Drehachse AS2-> GS_Position_und_Geschwindigkeit vorgeben"   // T42
      := "POS3_0_Signal"."-1001T1 Oriental_Positionen".POS_OK_Position[1];
   END_TRANSITION
   STEP Drehachse_GS:   // S40, max time T#10S, warning time T#7S
      supervision V := #Drehachse_GS.U > #Drehachse_GS.T_MAX;
              N    "POS3_0_Signal"."-1002T1 Oriental_Positionen".Start_POS_Position[1]
   END_STEP
   TRANSITION "T_Drehachse GS_2" FROM Drehachse_GS TO "Steckzyklus +1"   // T43
      := "POS3_0_Signal"."-1002T1 Oriental_Positionen".POS_OK_Position[1];
   END_TRANSITION
   STEP "Drehachse GS_auf_Absolut_0°_Richten":   // S41, max time T#10S, warning time T#7S
      supervision V := #"Drehachse GS_auf_Absolut_0°_Richten".U > #"Drehachse GS_auf_Absolut_0°_Richten".T_MAX;
              N    "POS3_0_Signal"."-1002T1 Oriental_Positionen".Start_POS_Position[1]
   END_STEP
   TRANSITION "T_Drehachse AS_2_Richten" FROM "Drehachse GS_auf_Absolut_0°_Richten" TO "Positionierachse GS_Richten_Position_und_Geschwindigkeit vorgeben"   // T44
      := "POS3_0_Signal"."-1002T1 Oriental_Positionen".POS_OK_Position[1];
   END_TRANSITION
   STEP "Wegmessung_Ausgleichszylinder in GS":   // S42, max time T#10S, warning time T#7S
      supervision V := #"Wegmessung_Ausgleichszylinder in GS".U > #"Wegmessung_Ausgleichszylinder in GS".T_MAX;
          S1  S    "POS3_0_Signal"."-POS3.0_Wegmessung_Ausgleichszylinder_Position_GS_aktiv"
          S1  R    "POS3_0_Signal"."-POS3.0_Wegmessung_Ausgleichszylinder_Position_AS1_aktiv"
          S1  N    "POS3_0_Signal"."-POS3.0_Wegmessung_Ausgleichszylinder_Sollwert_in_mm" := "Verwaltung_Teiledaten"."Wegmessung_Ausgleichszylinder Position GS"
          S1  R    "POS3_0_Signal".Status_gesteckt
   END_STEP
   TRANSITION "T_Wegmessung_Ausgleichszylinder in GS" FROM "Wegmessung_Ausgleichszylinder in GS" TO "Positionierachse GS_Position_und_Geschwindigkeit vorgeben"   // T45
      := "POS3_0_Signal"."-POS3.0_Wegmessung_Ausgleichszylinder_Position_GS_Abweichung_OK";
   END_TRANSITION
   STEP "Regelventil_Überlastzylinder  Sollwert":   // S44, max time T#10S, warning time T#7S
      supervision V := #"Regelventil_Überlastzylinder  Sollwert".U > #"Regelventil_Überlastzylinder  Sollwert".T_MAX;
          S1  N    "POS3_0_Signal"."-POS3_0_Regelventil_Überlastzylinder_Sollwert" := "Verwaltung_Teiledaten"."Druck p2 Überlastzylinder"
   END_STEP
   TRANSITION "T_Regelventil_Überlastzylinder  Sollwert" FROM "Regelventil_Überlastzylinder  Sollwert" TO "Positionierachse AS_Position_und_Geschwindigkeit vorgeben"   // T47
      := "POS3_0_Signal"."-POS3_0_Regelventil_Überlastzylinder_Abweichung_OK";
   END_TRANSITION
   STEP "Drehachse AS1_Position_und_Geschwindigkeit vorgeben":   // S37, max time T#10S, warning time T#7S
      supervision V := #"Drehachse AS1_Position_und_Geschwindigkeit vorgeben".U > #"Drehachse AS1_Position_und_Geschwindigkeit vorgeben".T_MAX;
          S1  N    "POS3_0_Signal"."-1002T1 Oriental_Positionen".Geschwindigkeit[2] := "Verwaltung_Teiledaten"."Drehantrieb Geschwindigkeit GS->AS1" / 6
          S1  N    "POS3_0_Signal"."-1002T1 Oriental_Positionen".Soll_Position[2] := "Verwaltung_Teiledaten"."Drehantrieb Position AS1"
   END_STEP
   TRANSITION "T_Drehachse AS1_Geschwindigkeit vorgeben" FROM "Drehachse AS1_Position_und_Geschwindigkeit vorgeben" TO "Drehachse AS1"   // T40
      := TRUE;
   END_TRANSITION
   STEP "Drehachse AS1-> GS_Position_und_Geschwindigkeit vorgeben":   // S38, max time T#10S, warning time T#7S
      supervision V := #"Drehachse AS1-> GS_Position_und_Geschwindigkeit vorgeben".U > #"Drehachse AS1-> GS_Position_und_Geschwindigkeit vorgeben".T_MAX;
          S1  N    "POS3_0_Signal"."-1002T1 Oriental_Positionen".Geschwindigkeit[3] := "Verwaltung_Teiledaten"."Drehantrieb Geschwindigkeit AS1->GS" / 6
          S1  N    "POS3_0_Signal"."-1002T1 Oriental_Positionen".Soll_Position[3] := 0.0 - "Verwaltung_Teiledaten"."Drehantrieb Position AS1"
   END_STEP
   TRANSITION "T_Drehachse AS1-> GS_Geschwindigkeit vorgeben" FROM "Drehachse AS1-> GS_Position_und_Geschwindigkeit vorgeben" TO "Drehachse GS"   // T41
      := TRUE;
   END_TRANSITION
   STEP "Regelventil_Ausgleichszylinder Sollwert":   // S43, max time T#10S, warning time T#7S
      supervision V := #"Regelventil_Ausgleichszylinder Sollwert".U > #"Regelventil_Ausgleichszylinder Sollwert".T_MAX;
          S1  N    "POS3_0_Signal"."-POS3_0_Regelventil_Ausgleichszylinder_Sollwert" := "Verwaltung_Teiledaten"."Druck p1 Ausgleichszylinder"
   END_STEP
   TRANSITION "T_Regelventil_Ausgleichszylinder Sollwert" FROM "Regelventil_Ausgleichszylinder Sollwert" TO "Regelventil_Überlastzylinder  Sollwert"   // T46
      := "POS3_0_Signal"."-POS3_0_Regelventil_Ausgleichszylinder_Abweichung_OK";
   END_TRANSITION
   STEP "Drehachse AS2-> GS_Position_und_Geschwindigkeit vorgeben":   // S45, max time T#10S, warning time T#7S
      supervision V := #"Drehachse AS2-> GS_Position_und_Geschwindigkeit vorgeben".U > #"Drehachse AS2-> GS_Position_und_Geschwindigkeit vorgeben".T_MAX;
          S1  N    "POS3_0_Signal"."-1002T1 Oriental_Positionen".Geschwindigkeit[1] := "Verwaltung_Teiledaten"."Drehantrieb Motorstrombegrenzung" / 6
          S1  N    "POS3_0_Signal"."-1002T1 Oriental_Positionen".Soll_Position[1] := "Verwaltung_Teiledaten"."Drehantrieb Position GS"
   END_STEP
   TRANSITION "T_Drehachse AS2-> GS_Geschwindigkeit vorgeben" FROM "Drehachse AS2-> GS_Position_und_Geschwindigkeit vorgeben" TO Drehachse_GS   // T48
      := TRUE;
   END_TRANSITION
   STEP "Positionierachse AS_Position_und_Geschwindigkeit vorgeben":   // S48, max time T#10S, warning time T#7S
      supervision V := #"Positionierachse AS_Position_und_Geschwindigkeit vorgeben".U > #"Positionierachse AS_Position_und_Geschwindigkeit vorgeben".T_MAX;
          S1  N    "POS3_0_Signal"."-1001T1 Oriental_Positionen".Geschwindigkeit[2] := "Verwaltung_Teiledaten"."Achse Geschwindigkeit GS->AS" / 150
          S1  N    "POS3_0_Signal"."-1001T1 Oriental_Positionen".Soll_Position[2] := "Verwaltung_Teiledaten"."Achse Position AS"
   END_STEP
   TRANSITION "T_Positionierachse AS_Position_und_Geschwindigkeit vorgeben" FROM "Positionierachse AS_Position_und_Geschwindigkeit vorgeben" TO "Positionierachse AS"   // T52
      := TRUE;
   END_TRANSITION
   STEP "Positionierachse GS_Position_und_Geschwindigkeit vorgeben":   // S49, max time T#10S, warning time T#7S
      supervision V := #"Positionierachse GS_Position_und_Geschwindigkeit vorgeben".U > #"Positionierachse GS_Position_und_Geschwindigkeit vorgeben".T_MAX;
          S1  N    "POS3_0_Signal"."-1001T1 Oriental_Positionen".Geschwindigkeit[1] := "Verwaltung_Teiledaten"."Achse Geschwindigkeit AS->GS" / 150
          S1  N    "POS3_0_Signal"."-1001T1 Oriental_Positionen".Soll_Position[1] := "Verwaltung_Teiledaten"."Achse Position GS"
   END_STEP
   TRANSITION "T_Positionierachse GS_Position_und_Geschwindigkeit vorgeben" FROM "Positionierachse GS_Position_und_Geschwindigkeit vorgeben" TO "Positionierachse GS"   // T53
      := TRUE;
   END_TRANSITION
   STEP "Positionierachse GS_Richten_Position_und_Geschwindigkeit vorgeben":   // S50, max time T#10S, warning time T#7S
      supervision V := #"Positionierachse GS_Richten_Position_und_Geschwindigkeit vorgeben".U > #"Positionierachse GS_Richten_Position_und_Geschwindigkeit vorgeben".T_MAX;
          S1  N    "POS3_0_Signal"."-1001T1 Oriental_Positionen".Geschwindigkeit[1] := 10.0
          S1  N    "POS3_0_Signal"."-1001T1 Oriental_Positionen".Soll_Position[1] := "Verwaltung_Teiledaten"."Achse Position GS"
   END_STEP
   TRANSITION "T_Positionierachse GS_Position_und_Geschwindigkeit vorgeben_1" FROM "Positionierachse GS_Richten_Position_und_Geschwindigkeit vorgeben" TO "Positionierachse GS_Richten"   // T54
      := TRUE;
   END_TRANSITION
   STEP "Steckzyklus +1":   // S51, max time T#10S, warning time T#7S
          S1  N    "POS3_0_Signal".Istzyklen := "POS3_0_Signal".Istzyklen +1
   END_STEP
   TRANSITION Steckzyklen_nicht_fertig FROM "Steckzyklus +1" TO Fertigmeldung   // T55
      := "POS3_0_Signal".Istzyklen < "POS3_0_Signal".Sollzyklen;
   END_TRANSITION
   TRANSITION Steckzyklen_fertig FROM "Steckzyklus +1" TO Automatikablauf_stoppen   // T64
      := "POS3_0_Signal".Istzyklen >= "POS3_0_Signal".Sollzyklen;
   END_TRANSITION
   STEP "Messmethode -- Messgerät ist bereit oder nicht verbunden":   // S56, max time T#10S, warning time T#7S
      supervision V := #"Messmethode -- Messgerät ist bereit oder nicht verbunden".U > T#30s;
   END_STEP
   TRANSITION T_Messmethode_AUS FROM "Messmethode -- Messgerät ist bereit oder nicht verbunden" TO "Regelventil_Ausgleichszylinder Sollwert"   // T3
      := "POS3_0_Signal".Kommunikation_Weiterschaltbedingungen_AUS;
   END_TRANSITION
   TRANSITION T_Messmethode_SP7_LabView FROM "Messmethode -- Messgerät ist bereit oder nicht verbunden" TO Messmethode_SP7_LabView_Messgerät_bereit_und_verbunden   // T66
      := "POS3_0_Signal".Kommunikation_Weiterschaltbedingungen_SP7;
   END_TRANSITION
   TRANSITION T_Messmethode_Digital FROM "Messmethode -- Messgerät ist bereit oder nicht verbunden" TO Messmethode_DIGITAL_Messgerät_bereit_und_verbunden   // T68
      := "POS3_0_Signal".Kommunikation_Weiterschaltbedingungen_DIGITAL;
   END_TRANSITION
   STEP "Position Drehachse abfragen":   // S57, max time T#10S, warning time T#7S
   END_STEP
   TRANSITION "T_Drehachse_kleiner_360°_und_größer_0°" FROM "Position Drehachse abfragen" TO "Drehachse GS_auf_Absolut_0°_Richten"   // T49
      := ("POS3_0_Signal"."-1002T1 Oriental_Absolute_Position" < 360.0) AND ("POS3_0_Signal"."-1002T1 Oriental_Absolute_Position" >= 0.0);
   END_TRANSITION
   TRANSITION "T_Drehachse_größer_360°_oder_kleiner_0°" FROM "Position Drehachse abfragen" TO "Drehachse AS1-> GS_Position_und_Geschwindigkeit vorgeben_Richten"   // T62
      := ("POS3_0_Signal"."-1002T1 Oriental_Absolute_Position" >= 360.0) OR ("POS3_0_Signal"."-1002T1 Oriental_Absolute_Position" < 0.0);
   END_TRANSITION
   STEP "Drehachse AS1-> GS_Richten":   // S47, max time T#10S, warning time T#7S
      supervision V := #"Drehachse AS1-> GS_Richten".U > #"Drehachse AS1-> GS_Richten".T_MAX;
              N    "POS3_0_Signal"."-1002T1 Oriental_Positionen".Start_POS_Position[3]
   END_STEP
   TRANSITION "T_Drehachse GS_1" FROM "Drehachse AS1-> GS_Richten" TO "Drehachse GS_auf_Absolut_0°_Richten"   // T51
      := "POS3_0_Signal"."-1002T1 Oriental_Positionen".POS_OK_Position[3];
   END_TRANSITION
   STEP "Drehachse AS1-> GS_Position_und_Geschwindigkeit vorgeben_Richten":   // S58, max time T#10S, warning time T#7S
      supervision V := #"Drehachse AS1-> GS_Position_und_Geschwindigkeit vorgeben_Richten".U > #"Drehachse AS1-> GS_Position_und_Geschwindigkeit vorgeben_Richten".T_MAX;
          S1  N    "POS3_0_Signal"."-1002T1 Oriental_Positionen".Geschwindigkeit[3] := "Verwaltung_Teiledaten"."Drehantrieb Geschwindigkeit AS1->GS" / 6
          S1  N    "POS3_0_Signal"."-1002T1 Oriental_Positionen".Soll_Position[3] := 0.0 - "POS3_0_Signal"."-1002T1 Oriental_Absolute_Position"
   END_STEP
   TRANSITION "T_Drehachse AS1-> GS_Geschwindigkeit vorgeben_Richten" FROM "Drehachse AS1-> GS_Position_und_Geschwindigkeit vorgeben_Richten" TO "Drehachse AS1-> GS_Richten"   // T63
      := #"Drehachse AS1-> GS_Position_und_Geschwindigkeit vorgeben_Richten".T > t#100MS;
   END_TRANSITION
   STEP Automatikablauf_stoppen:   // S59, max time T#10S, warning time T#7S
          S1  R    "HMI_Signale".Stop_nach_Zyklus
   END_STEP
   TRANSITION T_Automatikablauf_stoppen FROM Automatikablauf_stoppen TO Fertigmeldung   // T65
      := #Automatikablauf_stoppen.T > t#100MS;
   END_TRANSITION
   STEP Messmethode_SP7_LabView_Messgerät_bereit_und_verbunden:   // S60, max time T#10S, warning time T#7S
   END_STEP
   TRANSITION T_Messmethode_SP7_LabView_Messgerät_bereit_und_verbunden FROM Messmethode_SP7_LabView_Messgerät_bereit_und_verbunden TO "Regelventil_Ausgleichszylinder Sollwert"   // T67
      := "DB020_Com LabView"."E_Messgerät ist bereit und verbunden";
   END_TRANSITION
   STEP Messmethode_DIGITAL_Messgerät_bereit_und_verbunden:   // S61, max time T#10S, warning time T#7S
   END_STEP
   TRANSITION T_Messmethode_DIGITAL_Messgerät_bereit_und_verbunden FROM Messmethode_DIGITAL_Messgerät_bereit_und_verbunden TO "Regelventil_Ausgleichszylinder Sollwert"   // T69
      := false;
   END_TRANSITION
   STEP "Messmethode -- Startfreigabe Zwischenbefundung":   // S62, max time T#10S, warning time T#7S
   END_STEP
   TRANSITION "T_Messmethode_AUS -- Zwischenbefundung" FROM "Messmethode -- Startfreigabe Zwischenbefundung" TO "Wartezeit - Messmethode_AUS"   // T4
      := "POS3_0_Signal".Kommunikation_Weiterschaltbedingungen_AUS;
   END_TRANSITION
   TRANSITION "T_Messmethode_SP7_LabView -- Zwischenbefundung" FROM "Messmethode -- Startfreigabe Zwischenbefundung" TO "Wartezeit - Messmethode_SP7_LabView"   // T71
      := "POS3_0_Signal".Kommunikation_Weiterschaltbedingungen_SP7;
   END_TRANSITION
   TRANSITION "T_Messmethode_Digital -- Zwischenbefundung" FROM "Messmethode -- Startfreigabe Zwischenbefundung" TO "Wartezeit - Messmethode_Digital"   // T72
      := "POS3_0_Signal".Kommunikation_Weiterschaltbedingungen_DIGITAL;
   END_TRANSITION
   STEP "Wartezeit - Messmethode_SP7_LabView":   // S46, max time T#10S, warning time T#7S
          S1  S    "DB020_Com LabView".A_Startfreigabe_Zwischenbefundung
   END_STEP
   TRANSITION "T_Wartezeit abgelaufen - Messmethode_SP7_LabView" FROM "Wartezeit - Messmethode_SP7_LabView" TO "Rückmeldung_Startfreigabe_Zwischenbefundung_erhalten - Messmethode_SP7_LabView"   // T50
      := #"Wartezeit - Messmethode_SP7_LabView".T > "POS3_0_Signal"."Wartezeit Soll gesteckt";
   END_TRANSITION
   STEP "Zwischenbefundung ist fertig  - Messmethode_SP7_LabView":   // S63, max time T#10S, warning time T#7S
      supervision V := #"Zwischenbefundung ist fertig  - Messmethode_SP7_LabView".U > T#30s;
          S1  R    "DB020_Com LabView".A_Startfreigabe_Zwischenbefundung
   END_STEP
   TRANSITION "T_Zwischenbefundung ist fertig  - Messmethode_SP7_LabView" FROM "Zwischenbefundung ist fertig  - Messmethode_SP7_LabView" TO "Rückmeldung_Signal_Zwischenbfundung_erhalten  - Messmethode_SP7_LabView"   // T70
      := "DB020_Com LabView".E_Rückmeldung_Zwischenbefundung_fertig;
   END_TRANSITION
   STEP "Rückmeldung_Startfreigabe_Zwischenbefundung_erhalten - Messmethode_SP7_LabView":   // S64, max time T#10S, warning time T#7S
      supervision V := #"Rückmeldung_Startfreigabe_Zwischenbefundung_erhalten - Messmethode_SP7_LabView".U > t#30s;
   END_STEP
   TRANSITION "T_Zwischenbefudung ist gestartet  - Messmethode_SP7_LabView" FROM "Rückmeldung_Startfreigabe_Zwischenbefundung_erhalten - Messmethode_SP7_LabView" TO "Zwischenbefundung ist fertig  - Messmethode_SP7_LabView"   // T73
      := "DB020_Com LabView".E_Rückmeldung_Startfreigabe_Zwischenbefundung_erhalten;
   END_TRANSITION
   STEP "Rückmeldung_Signal_Zwischenbfundung_erhalten  - Messmethode_SP7_LabView":   // S65, max time T#10S, warning time T#7S
      supervision V := #"Rückmeldung_Signal_Zwischenbfundung_erhalten  - Messmethode_SP7_LabView".U > t#30S;
          S1  S    "DB020_Com LabView".A_Rückmeldung_Signal_Zwischenbfundung_erhalten
   END_STEP
   TRANSITION "T_Rückmeldung_Signal_Zwischenbfundung_erhalten  - Messmethode_SP7_LabView" FROM "Rückmeldung_Signal_Zwischenbfundung_erhalten  - Messmethode_SP7_LabView" TO "Rücksetzen Signale  - Messmethode_SP7_LabView"   // T74
      := NOT "DB020_Com LabView".E_Rückmeldung_Startfreigabe_Zwischenbefundung_erhalten AND NOT "DB020_Com LabView".E_Rückmeldung_Zwischenbefundung_fertig;
   END_TRANSITION
   STEP "Rücksetzen Signale  - Messmethode_SP7_LabView":   // S66, max time T#10S, warning time T#7S
      supervision V := #"Rücksetzen Signale  - Messmethode_SP7_LabView".U > t#30S;
          S1  R    "DB020_Com LabView".A_Rückmeldung_Signal_Zwischenbfundung_erhalten
          S1  R    "DB020_Com LabView".A_Startfreigabe_Zwischenbefundung
   END_STEP
   TRANSITION "T_Rücksetzen Signale  - Messmethode_SP7_LabView" FROM "Rücksetzen Signale  - Messmethode_SP7_LabView" TO "Drehachse AS1-> GS_Position_und_Geschwindigkeit vorgeben"   // T75
      := NOT "DB020_Com LabView".A_Rückmeldung_Signal_Zwischenbfundung_erhalten AND NOT "DB020_Com LabView".A_Startfreigabe_Zwischenbefundung;
   END_TRANSITION
   STEP "Wartezeit - Messmethode_Digital":   // S67, max time T#10S, warning time T#7S
   END_STEP
   TRANSITION "T_Wartezeit abgelaufen - Messmethode_Digital" FROM "Wartezeit - Messmethode_Digital" TO "Rückmeldung_Startfreigabe_Zwischenbefundung_erhalten - Messmethode_Digital"   // T76
      := #"Wartezeit - Messmethode_Digital".T > "POS3_0_Signal"."Wartezeit Soll gesteckt";
   END_TRANSITION
   STEP "Zwischenbefundung ist fertig  - Messmethode_Digital":   // S68, max time T#10S, warning time T#7S
      supervision V := #"Zwischenbefundung ist fertig  - Messmethode_Digital".U > T#30s;
   END_STEP
   TRANSITION "T_Zwischenbefundung ist fertig  - Messmethode_Digital" FROM "Zwischenbefundung ist fertig  - Messmethode_Digital" TO "Rückmeldung_Signal_Zwischenbfundung_erhalten - Messmethode_Digital"   // T77
      := false;
   END_TRANSITION
   STEP "Rückmeldung_Startfreigabe_Zwischenbefundung_erhalten - Messmethode_Digital":   // S69, max time T#10S, warning time T#7S
      supervision V := #"Rückmeldung_Startfreigabe_Zwischenbefundung_erhalten - Messmethode_Digital".U > t#30s;
   END_STEP
   TRANSITION "T_Zwischenbefudung ist gestartet - Messmethode_Digital" FROM "Rückmeldung_Startfreigabe_Zwischenbefundung_erhalten - Messmethode_Digital" TO "Zwischenbefundung ist fertig  - Messmethode_Digital"   // T78
      := false;
   END_TRANSITION
   STEP "Rückmeldung_Signal_Zwischenbfundung_erhalten - Messmethode_Digital":   // S70, max time T#10S, warning time T#7S
      supervision V := #"Rückmeldung_Signal_Zwischenbfundung_erhalten - Messmethode_Digital".U > t#30S;
   END_STEP
   TRANSITION "T_Rückmeldung_Signal_Zwischenbfundung_erhalten - Messmethode_Digital" FROM "Rückmeldung_Signal_Zwischenbfundung_erhalten - Messmethode_Digital" TO "Rücksetzen Signale  - Messmethode_Digital"   // T79
      := false;
   END_TRANSITION
   STEP "Rücksetzen Signale  - Messmethode_Digital":   // S71, max time T#10S, warning time T#7S
      supervision V := #"Rücksetzen Signale  - Messmethode_Digital".U > t#30S;
   END_STEP
   TRANSITION "T_Rücksetzen Signale  - Messmethode_Digital" FROM "Rücksetzen Signale  - Messmethode_Digital" TO "Drehachse AS1-> GS_Position_und_Geschwindigkeit vorgeben"   // T80
      := false;
   END_TRANSITION
END_FUNCTION_BLOCK

FUNCTION_BLOCK "Zaehler_Sicherheit"   // FB162, FBD
{ S7_Optimized_Access := 'TRUE' }
// stored: IsRetainMemResEnabled true, MemoryReserve 100, RetainMemoryReserve 100, SetENOAutomatically false
   VAR RETAIN
      "QS_NOT-HALT_Schuetz" { S7_SetPoint := 'True'} : CTU_UDINT;
      "QS_NOT-HALT_Tuere_1_RST" { S7_SetPoint := 'True'} : CTU_UDINT;
      "QS_NOT-HALT_Tuere_1" { S7_SetPoint := 'True'} : CTU_UDINT;
      "QS_NOT-HALT_Tuere_2_RST" { S7_SetPoint := 'True'} : CTU_UDINT;
      "QS_NOT-HALT_Tuere_2" { S7_SetPoint := 'True'} : CTU_UDINT;
      "QS_NOT-HALT_Roboter" { S7_SetPoint := 'True'} : CTU_UDINT;
      QS_Sichere_Bewegung { S7_SetPoint := 'True'} : CTU_UDINT;
      QS_Zuhaltung_Freigeben { S7_SetPoint := 'True'} : CTU_UDINT;
   END_VAR
BEGIN

REGION Network 1: Not Halt
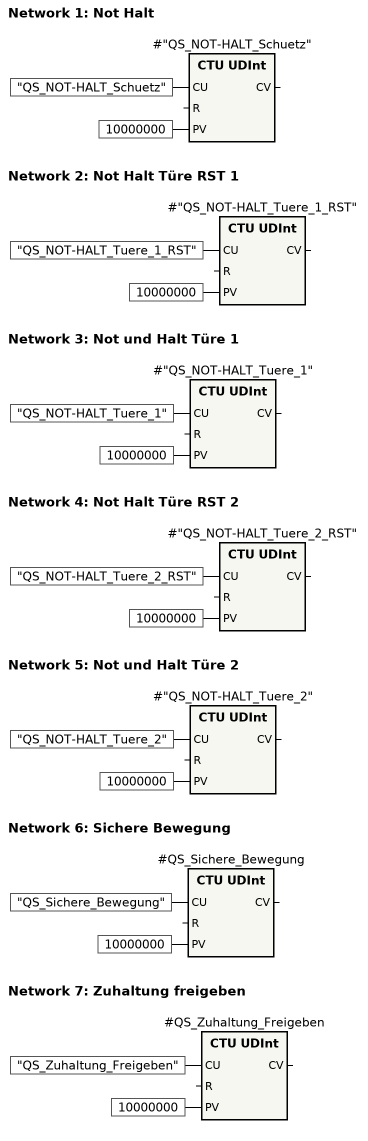
   #"QS_NOT-HALT_Schuetz"(CU := "QS_NOT-HALT_Schuetz", PV := 10000000);   // CTU
END_REGION

REGION Network 2: Not Halt Türe RST 1
   #"QS_NOT-HALT_Tuere_1_RST"(CU := "QS_NOT-HALT_Tuere_1_RST", PV := 10000000);   // CTU
END_REGION

REGION Network 3: Not und Halt Türe 1
   #"QS_NOT-HALT_Tuere_1"(CU := "QS_NOT-HALT_Tuere_1", PV := 10000000);   // CTU
END_REGION

REGION Network 4: Not Halt Türe RST 2
   #"QS_NOT-HALT_Tuere_2_RST"(CU := "QS_NOT-HALT_Tuere_2_RST", PV := 10000000);   // CTU
END_REGION

REGION Network 5: Not und Halt Türe 2
   #"QS_NOT-HALT_Tuere_2"(CU := "QS_NOT-HALT_Tuere_2", PV := 10000000);   // CTU
END_REGION

REGION Network 6: Sichere Bewegung
   #QS_Sichere_Bewegung(CU := "QS_Sichere_Bewegung", PV := 10000000);   // CTU
END_REGION

REGION Network 7: Zuhaltung freigeben
   #QS_Zuhaltung_Freigeben(CU := "QS_Zuhaltung_Freigeben", PV := 10000000);   // CTU
END_REGION
END_FUNCTION_BLOCK

FUNCTION_BLOCK "Main_Safety_RTG1"   // FB3, F_LAD
{ S7_Optimized_Access := 'TRUE' }
// stored: AutoNumber false
   VAR
      "ESTOP1_NOT-HALT Taster1" : ESTOP1;
      "stat_Q_NOT-HALT Taster1" : Bool;
      "stat_AckReq_NOT-HALT Taster1" : Bool;
      "ESTOP1_NOT-HALT Extern 1" : ESTOP1;
      "stat_Q_NOT-HALT Extern 1" : Bool;
      "stat_AckReq_NOT-HALT Extern1" : Bool;
      "ESTOP1_NOT-HALT Extern 2" : ESTOP1;
      "stat_Q_NOT-HALT Extern 2" : Bool;
      "stat_AckReq_NOT-HALT Extern 2" : Bool;
      "ESTOP1_Tür 1" : ESTOP1;
      "stat_Q_Tür 1" : Bool;
      "stat_AckReq_Tür 1" : Bool;
      "ESTOP1_Tür 2" : ESTOP1;
      "stat_Q_Tür 2" : Bool;
      "stat_AckReq_Tür 2" : Bool;
      ESTOP1_Systemdruck : ESTOP1;
      stat_AckReq_Systemdruck : Bool;
      "FDBACK_1_NOT-HALT Schütz mit DE_NOT-HALT_Schuetz_Rueckf" : FDBACK;
      "stat_Q_FDBK_1_NOT-HALT Schütz mit DE_NOT-HALT_Schuetz_Rueckf" : Bool;
      "stat_ERROR_FDBK_1_NOT-HALT Schütz mit DE_NOT-HALT_Schuetz_Rueckf" : Bool;
      "FDBACK_2_NOT-HALT Schütz mit IS_Rueck_Entlueftung" : FDBACK;
      "stat_Q_FDBK_2_NOT-HALT Schütz mit IS_Rueck_Entlueftung" : Bool;
      "stat_ERROR_FDBK_2_NOT-HALT Schütz mit IS_Rueck_Entlueftung" : Bool;
      "FDBACK_3_NOT-HALT Schütz mit IS_Druckbereich_entlueftet" : FDBACK;
      "stat_Q_FDBK_3_NOT-HALT Schütz mit IS_Druckbereich_entlueftet" : Bool;
      "stat_ERROR_FDBK_3_NOT-HALT Schütz mit IS_Druckbereich_entlueftet" : Bool;
      "FDBACK_4_NOT-HALT Türe 1 RST mit DE_NOT-HALT_Tuere_1_Rueck_RST" : FDBACK;
      "stat_Q_FDBK_4_NOT-HALT Türe 1 RST mit DE_NOT-HALT_Tuere_1_Rueck_RST" : Bool;
      "stat_ERROR_FDBK_4_NOT-HALT Türe 1 RST mit DE_NOT-HALT_Tuere_1_Rueck_RST" : Bool;
      "FDBACK_5_NOT-HALT Türe 1 mit DE_NOT-HALT_Tuere_1_Rueckf" : FDBACK;
      "stat_Q_FDBK_5_NOT-HALT Türe 1 mit DE_NOT-HALT_Tuere_1_Rueckf" : Bool;
      "stat_ERROR_FDBK_5_NOT-HALT Türe 1 mit DE_NOT-HALT_Tuere_1_Rueckf" : Bool;
      "FDBACK_6_NOT-HALT Türe 1 mit DE_Antriebe_Rueckf" : FDBACK;
      "stat_Q_FDBK_6_NOT-HALT Türe 1 mit DE_Antriebe_Rueckf" : Bool;
      "stat_ERROR_FDBK_6_NOT-HALT Türe 1 mit DE_Antriebe_Rueckf" : Bool;
      "FDBACK_7_NOT-HALT Türe 2 RST mit DE_NOT-HALT_Tuere_2_Rueck_RST" : FDBACK;
      "stat_Q_FDBK_7_NOT-HALT Türe 2 RST mit DE_NOT-HALT_Tuere_2_Rueck_RST" : Bool;
      "stat_ERROR_FDBK_7_NOT-HALT Türe 2 RST mit DE_NOT-HALT_Tuere_2_Rueck_RST" : Bool;
      "FDBACK_8_NOT-HALT Türe 2 mit DE_NOT-HALT_Tuere_2_Rueckf" : FDBACK;
      "stat_Q_FDBK_8_NOT-HALT Türe 2 mit DE_NOT-HALT_Tuere_2_Rueckf" : Bool;
      "stat_ERROR_FDBK_8_NOT-HALT Türe 2 mit DE_NOT-HALT_Tuere_2_Rueckf" : Bool;
      "FDBACK_10_Sicherere Bewegung" : FDBACK;
      "stat_AckReq_10_Sicherere Bewegung" : Bool;
      ACK_GL_Instance : ACK_GL;
      Systemdruck_OK : Bool;
      Antriebe_sicher : Bool;
      "TON_Zuhaltung_Freigben_mit_NOT-HALT" : TON;
      BA_0_groesser_1_5 : Bool;
      TON_BA_0_groesser_1_5 : TON;
      TON_Türen_setzen_zum_öffnen : TON;
      BA_0 : Bool;
      Zuhaltung_freigegeben : Bool;
   END_VAR
BEGIN

REGION Network 1: IS100_0/IS101_0 (2v2) NOT-HALT Taster 1
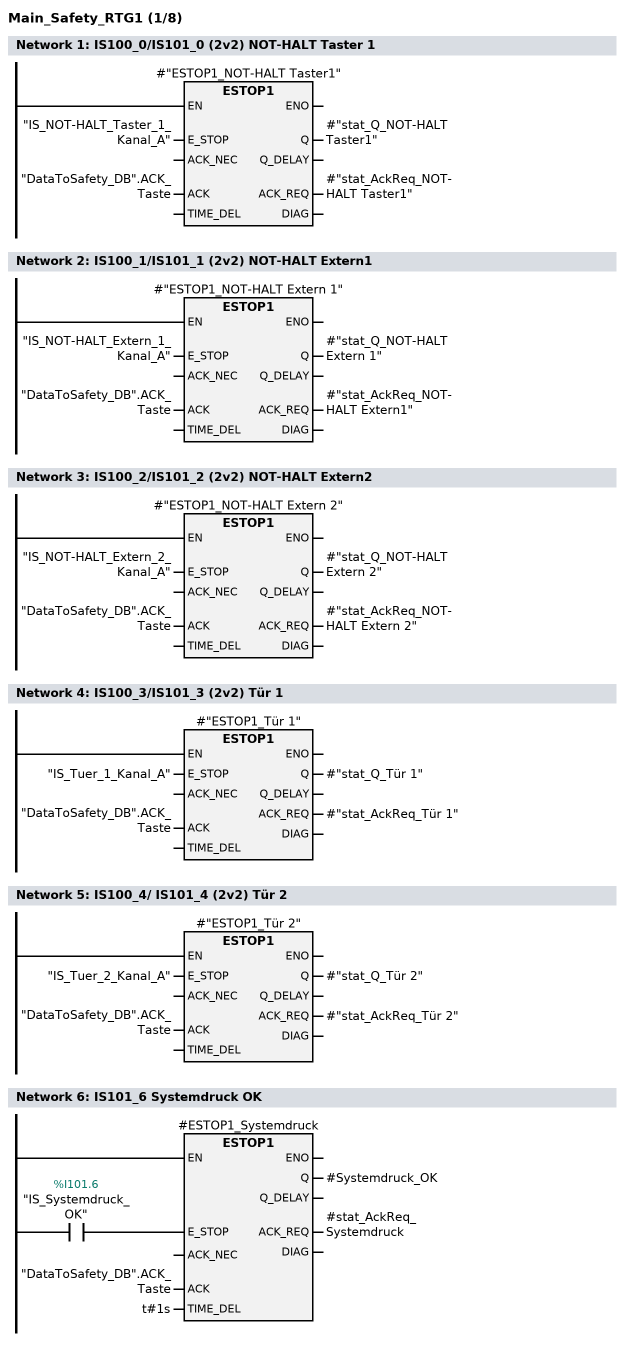
   RUNG wire#powerrail
      #"ESTOP1_NOT-HALT Taster1".ESTOP1(E_STOP := "IS_NOT-HALT_Taster_1_Kanal_A", ACK_NEC :=, ACK := "DataToSafety_DB".ACK_Taste, TIME_DEL :=, Q => #"stat_Q_NOT-HALT Taster1", Q_DELAY =>, ACK_REQ => #"stat_AckReq_NOT-HALT Taster1", DIAG =>)
   END_RUNG
   // the same network as SCL:
   #"ESTOP1_NOT-HALT Taster1"(E_STOP := "IS_NOT-HALT_Taster_1_Kanal_A",   // ESTOP1
                           ACK := "DataToSafety_DB".ACK_Taste,
                           Q => #"stat_Q_NOT-HALT Taster1",
                           ACK_REQ => #"stat_AckReq_NOT-HALT Taster1");
END_REGION

REGION Network 2: IS100_1/IS101_1 (2v2) NOT-HALT Extern1
   RUNG wire#powerrail
      #"ESTOP1_NOT-HALT Extern 1".ESTOP1(E_STOP := "IS_NOT-HALT_Extern_1_Kanal_A", ACK_NEC :=, ACK := "DataToSafety_DB".ACK_Taste, TIME_DEL :=, Q => #"stat_Q_NOT-HALT Extern 1", Q_DELAY =>, ACK_REQ => #"stat_AckReq_NOT-HALT Extern1", DIAG =>)
   END_RUNG
   // the same network as SCL:
   #"ESTOP1_NOT-HALT Extern 1"(E_STOP := "IS_NOT-HALT_Extern_1_Kanal_A",   // ESTOP1
                           ACK := "DataToSafety_DB".ACK_Taste,
                           Q => #"stat_Q_NOT-HALT Extern 1",
                           ACK_REQ => #"stat_AckReq_NOT-HALT Extern1");
END_REGION

REGION Network 3: IS100_2/IS101_2 (2v2) NOT-HALT Extern2
   RUNG wire#powerrail
      #"ESTOP1_NOT-HALT Extern 2".ESTOP1(E_STOP := "IS_NOT-HALT_Extern_2_Kanal_A", ACK_NEC :=, ACK := "DataToSafety_DB".ACK_Taste, TIME_DEL :=, Q => #"stat_Q_NOT-HALT Extern 2", Q_DELAY =>, ACK_REQ => #"stat_AckReq_NOT-HALT Extern 2", DIAG =>)
   END_RUNG
   // the same network as SCL:
   #"ESTOP1_NOT-HALT Extern 2"(E_STOP := "IS_NOT-HALT_Extern_2_Kanal_A",   // ESTOP1
                           ACK := "DataToSafety_DB".ACK_Taste,
                           Q => #"stat_Q_NOT-HALT Extern 2",
                           ACK_REQ => #"stat_AckReq_NOT-HALT Extern 2");
END_REGION

REGION Network 4: IS100_3/IS101_3 (2v2) Tür 1
   RUNG wire#powerrail
      #"ESTOP1_Tür 1".ESTOP1(E_STOP := "IS_Tuer_1_Kanal_A", ACK_NEC :=, ACK := "DataToSafety_DB".ACK_Taste, TIME_DEL :=, Q => #"stat_Q_Tür 1", Q_DELAY =>, ACK_REQ => #"stat_AckReq_Tür 1", DIAG =>)
   END_RUNG
   // the same network as SCL:
   #"ESTOP1_Tür 1"(E_STOP := "IS_Tuer_1_Kanal_A",   // ESTOP1
                   ACK := "DataToSafety_DB".ACK_Taste,
                   Q => #"stat_Q_Tür 1",
                   ACK_REQ => #"stat_AckReq_Tür 1");
END_REGION

REGION Network 5: IS100_4/ IS101_4 (2v2) Tür 2
   RUNG wire#powerrail
      #"ESTOP1_Tür 2".ESTOP1(E_STOP := "IS_Tuer_2_Kanal_A", ACK_NEC :=, ACK := "DataToSafety_DB".ACK_Taste, TIME_DEL :=, Q => #"stat_Q_Tür 2", Q_DELAY =>, ACK_REQ => #"stat_AckReq_Tür 2", DIAG =>)
   END_RUNG
   // the same network as SCL:
   #"ESTOP1_Tür 2"(E_STOP := "IS_Tuer_2_Kanal_A",   // ESTOP1
                   ACK := "DataToSafety_DB".ACK_Taste,
                   Q => #"stat_Q_Tür 2",
                   ACK_REQ => #"stat_AckReq_Tür 2");
END_REGION

REGION Network 6: IS101_6 Systemdruck OK
   RUNG wire#powerrail
      #ESTOP1_Systemdruck.ESTOP1(E_STOP := wire#w1, ACK_NEC :=, ACK := "DataToSafety_DB".ACK_Taste, TIME_DEL := t#1s, Q => #Systemdruck_OK, Q_DELAY =>, ACK_REQ => #stat_AckReq_Systemdruck, DIAG =>)
   END_RUNG
   RUNG wire#powerrail
      Contact( "IS_Systemdruck_OK" )
   END_RUNG wire#w1
   // the same network as SCL:
   #ESTOP1_Systemdruck(E_STOP := "IS_Systemdruck_OK",   // ESTOP1
                       ACK := "DataToSafety_DB".ACK_Taste,
                       TIME_DEL := t#1s,
                       Q => #Systemdruck_OK,
                       ACK_REQ => #stat_AckReq_Systemdruck);
END_REGION

REGION Network 7: Antriebe sicher
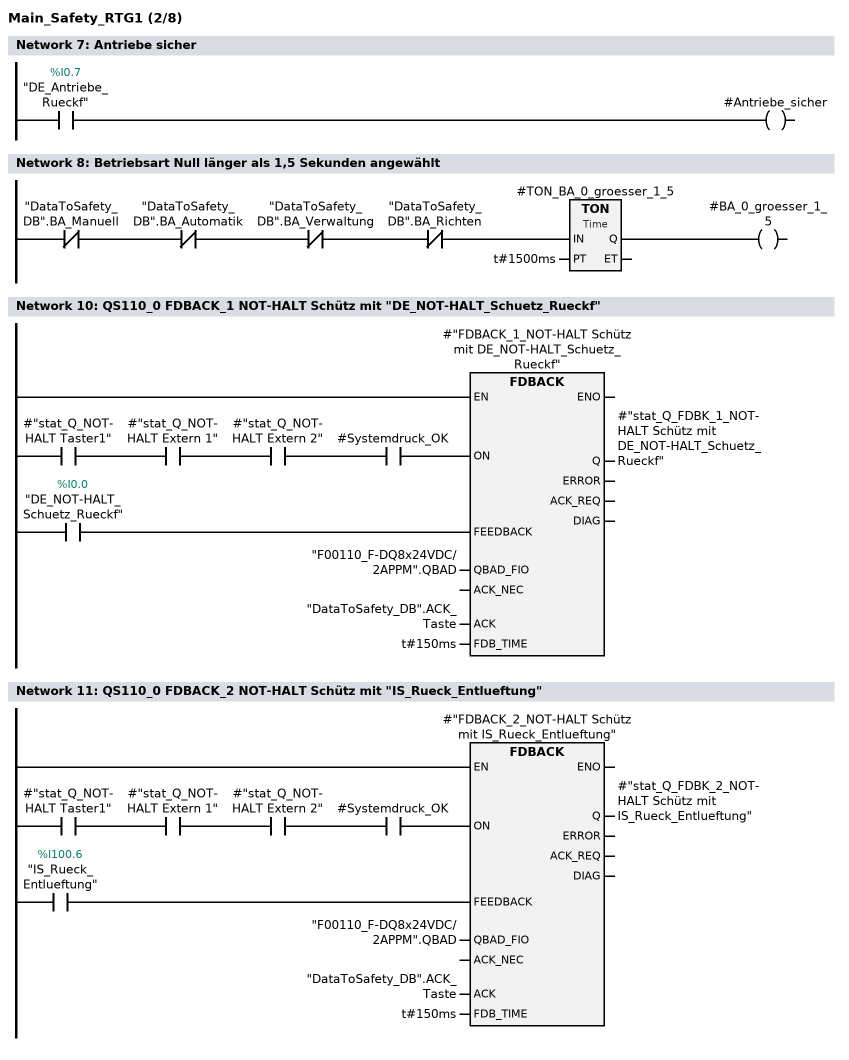
   RUNG wire#powerrail
      Contact( "DE_Antriebe_Rueckf" )
      Coil( #Antriebe_sicher )
   END_RUNG
   // the same network as SCL:
   #Antriebe_sicher := "DE_Antriebe_Rueckf";
END_REGION

REGION Network 8: Betriebsart Null länger als 1,5 Sekunden angewählt
   RUNG wire#powerrail
      I_Contact( "DataToSafety_DB".BA_Manuell )
      I_Contact( "DataToSafety_DB".BA_Automatik )
      I_Contact( "DataToSafety_DB".BA_Verwaltung )
      I_Contact( "DataToSafety_DB".BA_Richten )
      { S7_Templates := "[time_type := Time, codedbool_type := DInt]" } #TON_BA_0_groesser_1_5.TON(pt := t#1500ms, et =>)
      Coil( #BA_0_groesser_1_5 )
   END_RUNG
   // the same network as SCL:
   #TON_BA_0_groesser_1_5.TON(IN := NOT "DataToSafety_DB".BA_Manuell AND NOT "DataToSafety_DB".BA_Automatik AND NOT "DataToSafety_DB".BA_Verwaltung AND NOT "DataToSafety_DB".BA_Richten,
                           PT := t#1500ms);
   #BA_0_groesser_1_5 := #TON_BA_0_groesser_1_5.Q;
END_REGION

REGION Network 9: *********************************************************************************************
END_REGION

REGION Network 10: QS110_0 FDBACK_1 NOT-HALT Schütz mit "DE_NOT-HALT_Schuetz_Rueckf"
   RUNG wire#powerrail
      #"FDBACK_1_NOT-HALT Schütz mit DE_NOT-HALT_Schuetz_Rueckf".FDBACK(ON := wire#w1, FEEDBACK := wire#w2, QBAD_FIO := "F00110_F-DQ8x24VDC/2APPM".QBAD, ACK_NEC :=, ACK := "DataToSafety_DB".ACK_Taste, FDB_TIME := t#150ms, Q => #"stat_Q_FDBK_1_NOT-HALT Schütz mit DE_NOT-HALT_Schuetz_Rueckf", ERROR =>, ACK_REQ =>, DIAG =>)
   END_RUNG
   RUNG wire#powerrail
      Contact( #"stat_Q_NOT-HALT Taster1" )
      Contact( #"stat_Q_NOT-HALT Extern 1" )
      Contact( #"stat_Q_NOT-HALT Extern 2" )
      Contact( #Systemdruck_OK )
   END_RUNG wire#w1
   RUNG wire#powerrail
      Contact( "DE_NOT-HALT_Schuetz_Rueckf" )
   END_RUNG wire#w2
   // the same network as SCL:
   #"FDBACK_1_NOT-HALT Schütz mit DE_NOT-HALT_Schuetz_Rueckf"(ON := #"stat_Q_NOT-HALT Taster1" AND #"stat_Q_NOT-HALT Extern 1" AND #"stat_Q_NOT-HALT Extern 2" AND #Systemdruck_OK,   // FDBACK
                           FEEDBACK := "DE_NOT-HALT_Schuetz_Rueckf",
                           QBAD_FIO := "F00110_F-DQ8x24VDC/2APPM".QBAD,
                           ACK := "DataToSafety_DB".ACK_Taste,
                           FDB_TIME := t#150ms,
                           Q => #"stat_Q_FDBK_1_NOT-HALT Schütz mit DE_NOT-HALT_Schuetz_Rueckf");
END_REGION

REGION Network 11: QS110_0 FDBACK_2 NOT-HALT Schütz mit "IS_Rueck_Entlueftung"
   RUNG wire#powerrail
      #"FDBACK_2_NOT-HALT Schütz mit IS_Rueck_Entlueftung".FDBACK(ON := wire#w1, FEEDBACK := wire#w2, QBAD_FIO := "F00110_F-DQ8x24VDC/2APPM".QBAD, ACK_NEC :=, ACK := "DataToSafety_DB".ACK_Taste, FDB_TIME := t#150ms, Q => #"stat_Q_FDBK_2_NOT-HALT Schütz mit IS_Rueck_Entlueftung", ERROR =>, ACK_REQ =>, DIAG =>)
   END_RUNG
   RUNG wire#powerrail
      Contact( #"stat_Q_NOT-HALT Taster1" )
      Contact( #"stat_Q_NOT-HALT Extern 1" )
      Contact( #"stat_Q_NOT-HALT Extern 2" )
      Contact( #Systemdruck_OK )
   END_RUNG wire#w1
   RUNG wire#powerrail
      Contact( "IS_Rueck_Entlueftung" )
   END_RUNG wire#w2
   // the same network as SCL:
   #"FDBACK_2_NOT-HALT Schütz mit IS_Rueck_Entlueftung"(ON := #"stat_Q_NOT-HALT Taster1" AND #"stat_Q_NOT-HALT Extern 1" AND #"stat_Q_NOT-HALT Extern 2" AND #Systemdruck_OK,   // FDBACK
                           FEEDBACK := "IS_Rueck_Entlueftung",
                           QBAD_FIO := "F00110_F-DQ8x24VDC/2APPM".QBAD,
                           ACK := "DataToSafety_DB".ACK_Taste,
                           FDB_TIME := t#150ms,
                           Q => #"stat_Q_FDBK_2_NOT-HALT Schütz mit IS_Rueck_Entlueftung");
END_REGION

REGION Network 12: QS110_0 FDBACK_3 NOT-HALT Schütz mit "IS_Druckbereich_entlueftet"
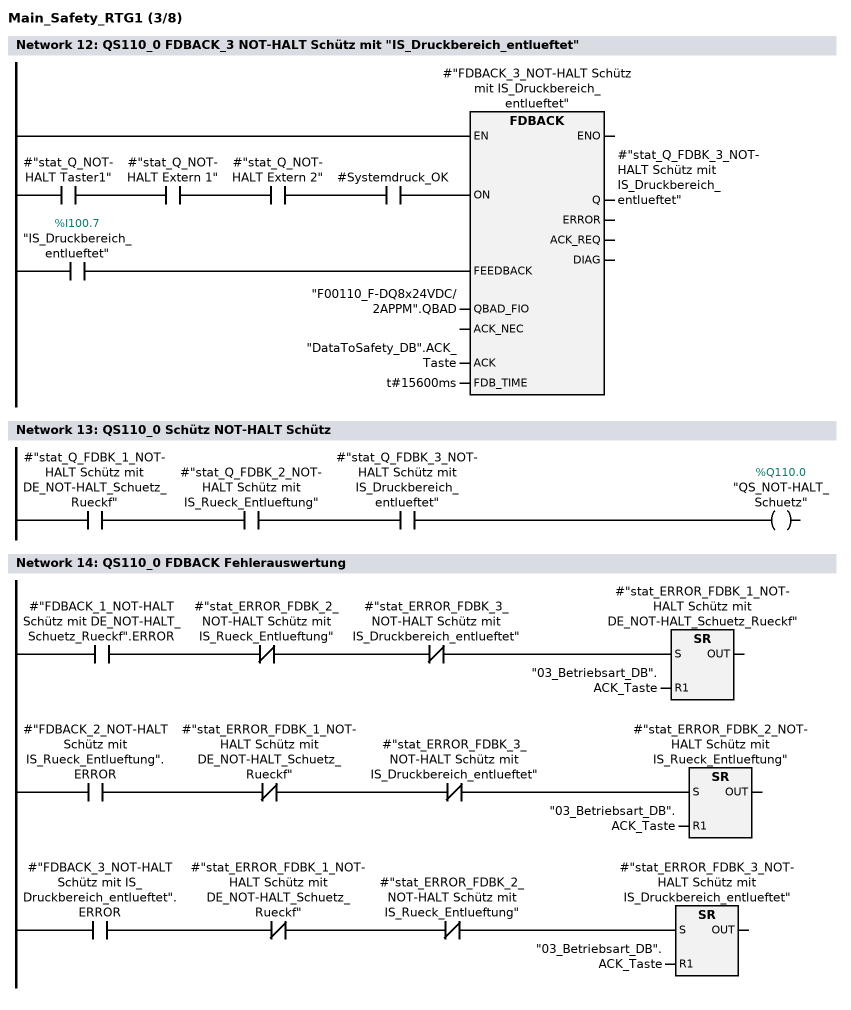
   RUNG wire#powerrail
      #"FDBACK_3_NOT-HALT Schütz mit IS_Druckbereich_entlueftet".FDBACK(ON := wire#w1, FEEDBACK := wire#w2, QBAD_FIO := "F00110_F-DQ8x24VDC/2APPM".QBAD, ACK_NEC :=, ACK := "DataToSafety_DB".ACK_Taste, FDB_TIME := t#15600ms, Q => #"stat_Q_FDBK_3_NOT-HALT Schütz mit IS_Druckbereich_entlueftet", ERROR =>, ACK_REQ =>, DIAG =>)
   END_RUNG
   RUNG wire#powerrail
      Contact( #"stat_Q_NOT-HALT Taster1" )
      Contact( #"stat_Q_NOT-HALT Extern 1" )
      Contact( #"stat_Q_NOT-HALT Extern 2" )
      Contact( #Systemdruck_OK )
   END_RUNG wire#w1
   RUNG wire#powerrail
      Contact( "IS_Druckbereich_entlueftet" )
   END_RUNG wire#w2
   // the same network as SCL:
   #"FDBACK_3_NOT-HALT Schütz mit IS_Druckbereich_entlueftet"(ON := #"stat_Q_NOT-HALT Taster1" AND #"stat_Q_NOT-HALT Extern 1" AND #"stat_Q_NOT-HALT Extern 2" AND #Systemdruck_OK,   // FDBACK
                           FEEDBACK := "IS_Druckbereich_entlueftet",
                           QBAD_FIO := "F00110_F-DQ8x24VDC/2APPM".QBAD,
                           ACK := "DataToSafety_DB".ACK_Taste,
                           FDB_TIME := t#15600ms,
                           Q => #"stat_Q_FDBK_3_NOT-HALT Schütz mit IS_Druckbereich_entlueftet");
END_REGION

REGION Network 13: QS110_0 Schütz NOT-HALT Schütz
   RUNG wire#powerrail
      Contact( #"stat_Q_FDBK_1_NOT-HALT Schütz mit DE_NOT-HALT_Schuetz_Rueckf" )
      Contact( #"stat_Q_FDBK_2_NOT-HALT Schütz mit IS_Rueck_Entlueftung" )
      Contact( #"stat_Q_FDBK_3_NOT-HALT Schütz mit IS_Druckbereich_entlueftet" )
      Coil( "QS_NOT-HALT_Schuetz" )
   END_RUNG
   // the same network as SCL:
   "QS_NOT-HALT_Schuetz" := #"stat_Q_FDBK_1_NOT-HALT Schütz mit DE_NOT-HALT_Schuetz_Rueckf" AND #"stat_Q_FDBK_2_NOT-HALT Schütz mit IS_Rueck_Entlueftung" AND #"stat_Q_FDBK_3_NOT-HALT Schütz mit IS_Druckbereich_entlueftet";
END_REGION

REGION Network 14: QS110_0 FDBACK Fehlerauswertung
   RUNG wire#powerrail
      Contact( #"FDBACK_1_NOT-HALT Schütz mit DE_NOT-HALT_Schuetz_Rueckf".ERROR )
      I_Contact( #"stat_ERROR_FDBK_2_NOT-HALT Schütz mit IS_Rueck_Entlueftung" )
      I_Contact( #"stat_ERROR_FDBK_3_NOT-HALT Schütz mit IS_Druckbereich_entlueftet" )
      S_SR(operand := #"stat_ERROR_FDBK_1_NOT-HALT Schütz mit DE_NOT-HALT_Schuetz_Rueckf", r1 := "03_Betriebsart_DB".ACK_Taste)
   END_RUNG
   RUNG wire#powerrail
      Contact( #"FDBACK_2_NOT-HALT Schütz mit IS_Rueck_Entlueftung".ERROR )
      I_Contact( #"stat_ERROR_FDBK_1_NOT-HALT Schütz mit DE_NOT-HALT_Schuetz_Rueckf" )
      I_Contact( #"stat_ERROR_FDBK_3_NOT-HALT Schütz mit IS_Druckbereich_entlueftet" )
      S_SR(operand := #"stat_ERROR_FDBK_2_NOT-HALT Schütz mit IS_Rueck_Entlueftung", r1 := "03_Betriebsart_DB".ACK_Taste)
   END_RUNG
   RUNG wire#powerrail
      Contact( #"FDBACK_3_NOT-HALT Schütz mit IS_Druckbereich_entlueftet".ERROR )
      I_Contact( #"stat_ERROR_FDBK_1_NOT-HALT Schütz mit DE_NOT-HALT_Schuetz_Rueckf" )
      I_Contact( #"stat_ERROR_FDBK_2_NOT-HALT Schütz mit IS_Rueck_Entlueftung" )
      S_SR(operand := #"stat_ERROR_FDBK_3_NOT-HALT Schütz mit IS_Druckbereich_entlueftet", r1 := "03_Betriebsart_DB".ACK_Taste)
   END_RUNG
   // the same network as SCL:
   IF #"FDBACK_1_NOT-HALT Schütz mit DE_NOT-HALT_Schuetz_Rueckf".ERROR AND NOT #"stat_ERROR_FDBK_2_NOT-HALT Schütz mit IS_Rueck_Entlueftung" AND NOT #"stat_ERROR_FDBK_3_NOT-HALT Schütz mit IS_Druckbereich_entlueftet" THEN
       #"stat_ERROR_FDBK_1_NOT-HALT Schütz mit DE_NOT-HALT_Schuetz_Rueckf" := TRUE;   // SR flip-flop
   END_IF;
   IF "03_Betriebsart_DB".ACK_Taste THEN
       #"stat_ERROR_FDBK_1_NOT-HALT Schütz mit DE_NOT-HALT_Schuetz_Rueckf" := FALSE;
   END_IF;
   IF #"FDBACK_2_NOT-HALT Schütz mit IS_Rueck_Entlueftung".ERROR AND NOT #"stat_ERROR_FDBK_1_NOT-HALT Schütz mit DE_NOT-HALT_Schuetz_Rueckf" AND NOT #"stat_ERROR_FDBK_3_NOT-HALT Schütz mit IS_Druckbereich_entlueftet" THEN
       #"stat_ERROR_FDBK_2_NOT-HALT Schütz mit IS_Rueck_Entlueftung" := TRUE;   // SR flip-flop
   END_IF;
   IF "03_Betriebsart_DB".ACK_Taste THEN
       #"stat_ERROR_FDBK_2_NOT-HALT Schütz mit IS_Rueck_Entlueftung" := FALSE;
   END_IF;
   IF #"FDBACK_3_NOT-HALT Schütz mit IS_Druckbereich_entlueftet".ERROR AND NOT #"stat_ERROR_FDBK_1_NOT-HALT Schütz mit DE_NOT-HALT_Schuetz_Rueckf" AND NOT #"stat_ERROR_FDBK_2_NOT-HALT Schütz mit IS_Rueck_Entlueftung" THEN
       #"stat_ERROR_FDBK_3_NOT-HALT Schütz mit IS_Druckbereich_entlueftet" := TRUE;   // SR flip-flop
   END_IF;
   IF "03_Betriebsart_DB".ACK_Taste THEN
       #"stat_ERROR_FDBK_3_NOT-HALT Schütz mit IS_Druckbereich_entlueftet" := FALSE;
   END_IF;
END_REGION

REGION Network 15: *********************************************************************************************
END_REGION

REGION Network 16: QS110_1 FDBACK_4 NOT-HALT Türe 1 RST mit "DE_NOT-HALT_Tuere_1_RST_Rueck"
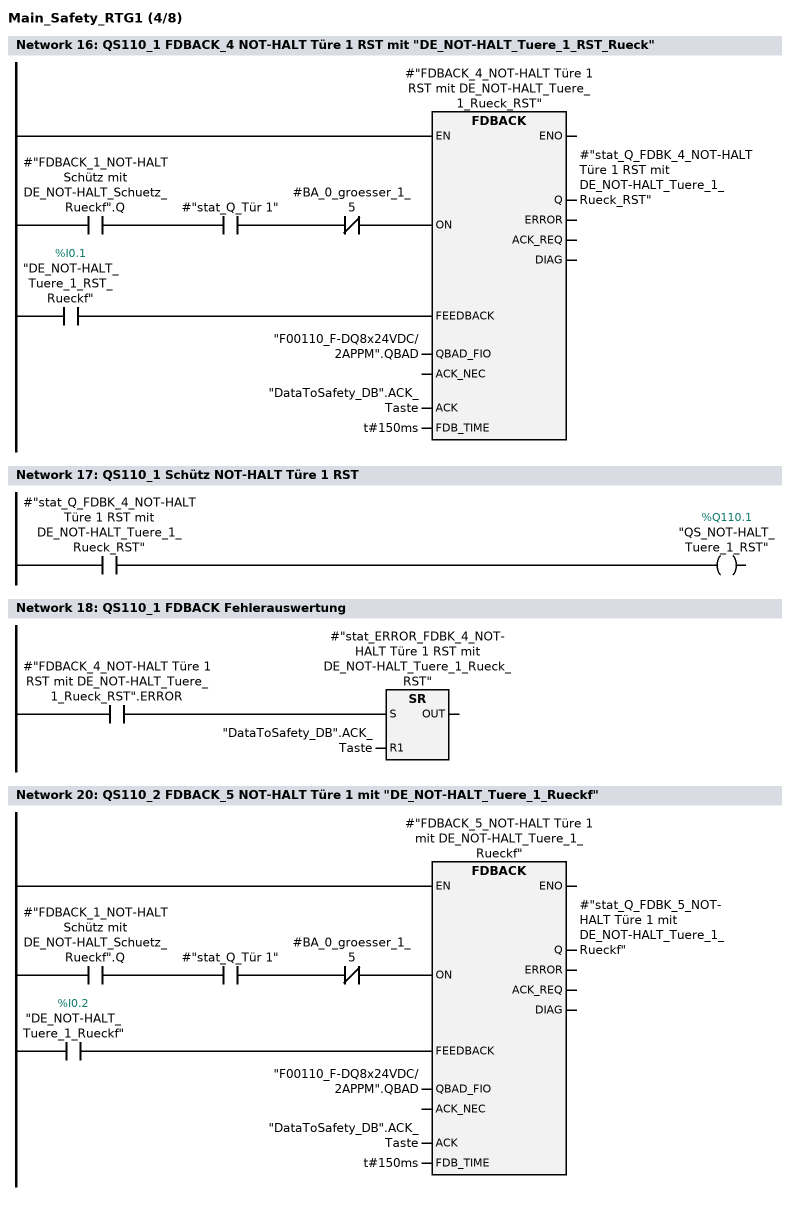
   RUNG wire#powerrail
      #"FDBACK_4_NOT-HALT Türe 1 RST mit DE_NOT-HALT_Tuere_1_Rueck_RST".FDBACK(ON := wire#w1, FEEDBACK := wire#w2, QBAD_FIO := "F00110_F-DQ8x24VDC/2APPM".QBAD, ACK_NEC :=, ACK := "DataToSafety_DB".ACK_Taste, FDB_TIME := t#150ms, Q => #"stat_Q_FDBK_4_NOT-HALT Türe 1 RST mit DE_NOT-HALT_Tuere_1_Rueck_RST", ERROR =>, ACK_REQ =>, DIAG =>)
   END_RUNG
   RUNG wire#powerrail
      Contact( #"FDBACK_1_NOT-HALT Schütz mit DE_NOT-HALT_Schuetz_Rueckf".Q )
      Contact( #"stat_Q_Tür 1" )
      I_Contact( #BA_0_groesser_1_5 )
   END_RUNG wire#w1
   RUNG wire#powerrail
      Contact( "DE_NOT-HALT_Tuere_1_RST_Rueckf" )
   END_RUNG wire#w2
   // the same network as SCL:
   #"FDBACK_4_NOT-HALT Türe 1 RST mit DE_NOT-HALT_Tuere_1_Rueck_RST"(ON := #"FDBACK_1_NOT-HALT Schütz mit DE_NOT-HALT_Schuetz_Rueckf".Q AND #"stat_Q_Tür 1" AND NOT #BA_0_groesser_1_5,   // FDBACK
                           FEEDBACK := "DE_NOT-HALT_Tuere_1_RST_Rueckf",
                           QBAD_FIO := "F00110_F-DQ8x24VDC/2APPM".QBAD,
                           ACK := "DataToSafety_DB".ACK_Taste,
                           FDB_TIME := t#150ms,
                           Q => #"stat_Q_FDBK_4_NOT-HALT Türe 1 RST mit DE_NOT-HALT_Tuere_1_Rueck_RST");
END_REGION

REGION Network 17: QS110_1 Schütz NOT-HALT Türe 1 RST
   RUNG wire#powerrail
      Contact( #"stat_Q_FDBK_4_NOT-HALT Türe 1 RST mit DE_NOT-HALT_Tuere_1_Rueck_RST" )
      Coil( "QS_NOT-HALT_Tuere_1_RST" )
   END_RUNG
   // the same network as SCL:
   "QS_NOT-HALT_Tuere_1_RST" := #"stat_Q_FDBK_4_NOT-HALT Türe 1 RST mit DE_NOT-HALT_Tuere_1_Rueck_RST";
END_REGION

REGION Network 18: QS110_1 FDBACK Fehlerauswertung
   RUNG wire#powerrail
      Contact( #"FDBACK_4_NOT-HALT Türe 1 RST mit DE_NOT-HALT_Tuere_1_Rueck_RST".ERROR )
      S_SR(operand := #"stat_ERROR_FDBK_4_NOT-HALT Türe 1 RST mit DE_NOT-HALT_Tuere_1_Rueck_RST", r1 := "DataToSafety_DB".ACK_Taste)
   END_RUNG
   // the same network as SCL:
   IF #"FDBACK_4_NOT-HALT Türe 1 RST mit DE_NOT-HALT_Tuere_1_Rueck_RST".ERROR THEN
       #"stat_ERROR_FDBK_4_NOT-HALT Türe 1 RST mit DE_NOT-HALT_Tuere_1_Rueck_RST" := TRUE;   // SR flip-flop
   END_IF;
   IF "DataToSafety_DB".ACK_Taste THEN
       #"stat_ERROR_FDBK_4_NOT-HALT Türe 1 RST mit DE_NOT-HALT_Tuere_1_Rueck_RST" := FALSE;
   END_IF;
END_REGION

REGION Network 19: *********************************************************************************************
END_REGION

REGION Network 20: QS110_2 FDBACK_5 NOT-HALT Türe 1 mit "DE_NOT-HALT_Tuere_1_Rueckf"
   RUNG wire#powerrail
      #"FDBACK_5_NOT-HALT Türe 1 mit DE_NOT-HALT_Tuere_1_Rueckf".FDBACK(ON := wire#w1, FEEDBACK := wire#w2, QBAD_FIO := "F00110_F-DQ8x24VDC/2APPM".QBAD, ACK_NEC :=, ACK := "DataToSafety_DB".ACK_Taste, FDB_TIME := t#150ms, Q => #"stat_Q_FDBK_5_NOT-HALT Türe 1 mit DE_NOT-HALT_Tuere_1_Rueckf", ERROR =>, ACK_REQ =>, DIAG =>)
   END_RUNG
   RUNG wire#powerrail
      Contact( #"FDBACK_1_NOT-HALT Schütz mit DE_NOT-HALT_Schuetz_Rueckf".Q )
      Contact( #"stat_Q_Tür 1" )
      I_Contact( #BA_0_groesser_1_5 )
   END_RUNG wire#w1
   RUNG wire#powerrail
      Contact( "DE_NOT-HALT_Tuere_1_Rueckf" )
   END_RUNG wire#w2
   // the same network as SCL:
   #"FDBACK_5_NOT-HALT Türe 1 mit DE_NOT-HALT_Tuere_1_Rueckf"(ON := #"FDBACK_1_NOT-HALT Schütz mit DE_NOT-HALT_Schuetz_Rueckf".Q AND #"stat_Q_Tür 1" AND NOT #BA_0_groesser_1_5,   // FDBACK
                           FEEDBACK := "DE_NOT-HALT_Tuere_1_Rueckf",
                           QBAD_FIO := "F00110_F-DQ8x24VDC/2APPM".QBAD,
                           ACK := "DataToSafety_DB".ACK_Taste,
                           FDB_TIME := t#150ms,
                           Q => #"stat_Q_FDBK_5_NOT-HALT Türe 1 mit DE_NOT-HALT_Tuere_1_Rueckf");
END_REGION

REGION Network 21: QS110_2 FDBACK_6 NOT-HALT Türe 1 mit "DE_Antriebe_Rueckf"
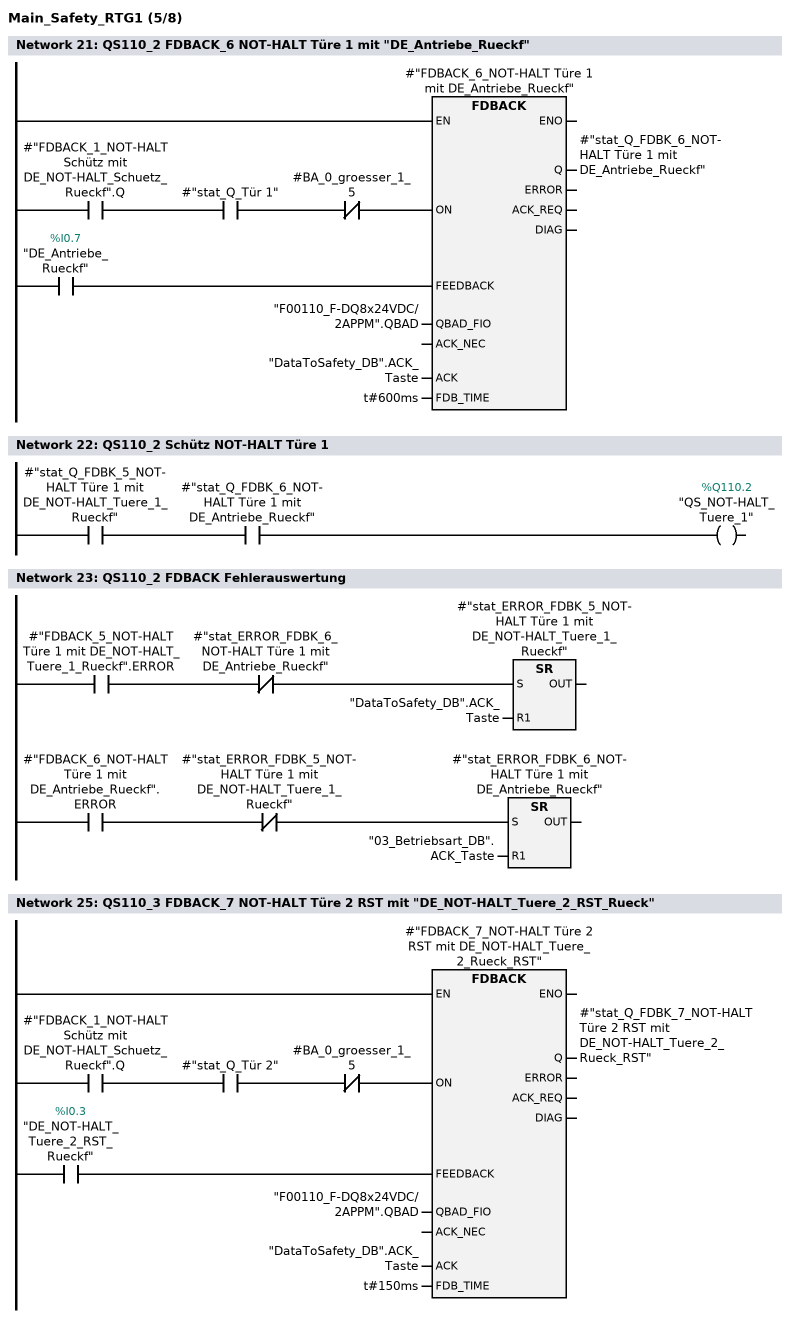
   RUNG wire#powerrail
      #"FDBACK_6_NOT-HALT Türe 1 mit DE_Antriebe_Rueckf".FDBACK(ON := wire#w1, FEEDBACK := wire#w2, QBAD_FIO := "F00110_F-DQ8x24VDC/2APPM".QBAD, ACK_NEC :=, ACK := "DataToSafety_DB".ACK_Taste, FDB_TIME := t#600ms, Q => #"stat_Q_FDBK_6_NOT-HALT Türe 1 mit DE_Antriebe_Rueckf", ERROR =>, ACK_REQ =>, DIAG =>)
   END_RUNG
   RUNG wire#powerrail
      Contact( #"FDBACK_1_NOT-HALT Schütz mit DE_NOT-HALT_Schuetz_Rueckf".Q )
      Contact( #"stat_Q_Tür 1" )
      I_Contact( #BA_0_groesser_1_5 )
   END_RUNG wire#w1
   RUNG wire#powerrail
      Contact( "DE_Antriebe_Rueckf" )
   END_RUNG wire#w2
   // the same network as SCL:
   #"FDBACK_6_NOT-HALT Türe 1 mit DE_Antriebe_Rueckf"(ON := #"FDBACK_1_NOT-HALT Schütz mit DE_NOT-HALT_Schuetz_Rueckf".Q AND #"stat_Q_Tür 1" AND NOT #BA_0_groesser_1_5,   // FDBACK
                           FEEDBACK := "DE_Antriebe_Rueckf",
                           QBAD_FIO := "F00110_F-DQ8x24VDC/2APPM".QBAD,
                           ACK := "DataToSafety_DB".ACK_Taste,
                           FDB_TIME := t#600ms,
                           Q => #"stat_Q_FDBK_6_NOT-HALT Türe 1 mit DE_Antriebe_Rueckf");
END_REGION

REGION Network 22: QS110_2 Schütz NOT-HALT Türe 1
   RUNG wire#powerrail
      Contact( #"stat_Q_FDBK_5_NOT-HALT Türe 1 mit DE_NOT-HALT_Tuere_1_Rueckf" )
      Contact( #"stat_Q_FDBK_6_NOT-HALT Türe 1 mit DE_Antriebe_Rueckf" )
      Coil( "QS_NOT-HALT_Tuere_1" )
   END_RUNG
   // the same network as SCL:
   "QS_NOT-HALT_Tuere_1" := #"stat_Q_FDBK_5_NOT-HALT Türe 1 mit DE_NOT-HALT_Tuere_1_Rueckf" AND #"stat_Q_FDBK_6_NOT-HALT Türe 1 mit DE_Antriebe_Rueckf";
END_REGION

REGION Network 23: QS110_2 FDBACK Fehlerauswertung
   RUNG wire#powerrail
      Contact( #"FDBACK_5_NOT-HALT Türe 1 mit DE_NOT-HALT_Tuere_1_Rueckf".ERROR )
      I_Contact( #"stat_ERROR_FDBK_6_NOT-HALT Türe 1 mit DE_Antriebe_Rueckf" )
      S_SR(operand := #"stat_ERROR_FDBK_5_NOT-HALT Türe 1 mit DE_NOT-HALT_Tuere_1_Rueckf", r1 := "DataToSafety_DB".ACK_Taste)
   END_RUNG
   RUNG wire#powerrail
      Contact( #"FDBACK_6_NOT-HALT Türe 1 mit DE_Antriebe_Rueckf".ERROR )
      I_Contact( #"stat_ERROR_FDBK_5_NOT-HALT Türe 1 mit DE_NOT-HALT_Tuere_1_Rueckf" )
      S_SR(operand := #"stat_ERROR_FDBK_6_NOT-HALT Türe 1 mit DE_Antriebe_Rueckf", r1 := "03_Betriebsart_DB".ACK_Taste)
   END_RUNG
   // the same network as SCL:
   IF #"FDBACK_5_NOT-HALT Türe 1 mit DE_NOT-HALT_Tuere_1_Rueckf".ERROR AND NOT #"stat_ERROR_FDBK_6_NOT-HALT Türe 1 mit DE_Antriebe_Rueckf" THEN
       #"stat_ERROR_FDBK_5_NOT-HALT Türe 1 mit DE_NOT-HALT_Tuere_1_Rueckf" := TRUE;   // SR flip-flop
   END_IF;
   IF "DataToSafety_DB".ACK_Taste THEN
       #"stat_ERROR_FDBK_5_NOT-HALT Türe 1 mit DE_NOT-HALT_Tuere_1_Rueckf" := FALSE;
   END_IF;
   IF #"FDBACK_6_NOT-HALT Türe 1 mit DE_Antriebe_Rueckf".ERROR AND NOT #"stat_ERROR_FDBK_5_NOT-HALT Türe 1 mit DE_NOT-HALT_Tuere_1_Rueckf" THEN
       #"stat_ERROR_FDBK_6_NOT-HALT Türe 1 mit DE_Antriebe_Rueckf" := TRUE;   // SR flip-flop
   END_IF;
   IF "03_Betriebsart_DB".ACK_Taste THEN
       #"stat_ERROR_FDBK_6_NOT-HALT Türe 1 mit DE_Antriebe_Rueckf" := FALSE;
   END_IF;
END_REGION

REGION Network 24: *********************************************************************************************
END_REGION

REGION Network 25: QS110_3 FDBACK_7 NOT-HALT Türe 2 RST mit "DE_NOT-HALT_Tuere_2_RST_Rueck"
   RUNG wire#powerrail
      #"FDBACK_7_NOT-HALT Türe 2 RST mit DE_NOT-HALT_Tuere_2_Rueck_RST".FDBACK(ON := wire#w1, FEEDBACK := wire#w2, QBAD_FIO := "F00110_F-DQ8x24VDC/2APPM".QBAD, ACK_NEC :=, ACK := "DataToSafety_DB".ACK_Taste, FDB_TIME := t#150ms, Q => #"stat_Q_FDBK_7_NOT-HALT Türe 2 RST mit DE_NOT-HALT_Tuere_2_Rueck_RST", ERROR =>, ACK_REQ =>, DIAG =>)
   END_RUNG
   RUNG wire#powerrail
      Contact( #"FDBACK_1_NOT-HALT Schütz mit DE_NOT-HALT_Schuetz_Rueckf".Q )
      Contact( #"stat_Q_Tür 2" )
      I_Contact( #BA_0_groesser_1_5 )
   END_RUNG wire#w1
   RUNG wire#powerrail
      Contact( "DE_NOT-HALT_Tuere_2_RST_Rueckf" )
   END_RUNG wire#w2
   // the same network as SCL:
   #"FDBACK_7_NOT-HALT Türe 2 RST mit DE_NOT-HALT_Tuere_2_Rueck_RST"(ON := #"FDBACK_1_NOT-HALT Schütz mit DE_NOT-HALT_Schuetz_Rueckf".Q AND #"stat_Q_Tür 2" AND NOT #BA_0_groesser_1_5,   // FDBACK
                           FEEDBACK := "DE_NOT-HALT_Tuere_2_RST_Rueckf",
                           QBAD_FIO := "F00110_F-DQ8x24VDC/2APPM".QBAD,
                           ACK := "DataToSafety_DB".ACK_Taste,
                           FDB_TIME := t#150ms,
                           Q => #"stat_Q_FDBK_7_NOT-HALT Türe 2 RST mit DE_NOT-HALT_Tuere_2_Rueck_RST");
END_REGION

REGION Network 26: QS110_3 Schütz NOT-HALT Türe 2 RST
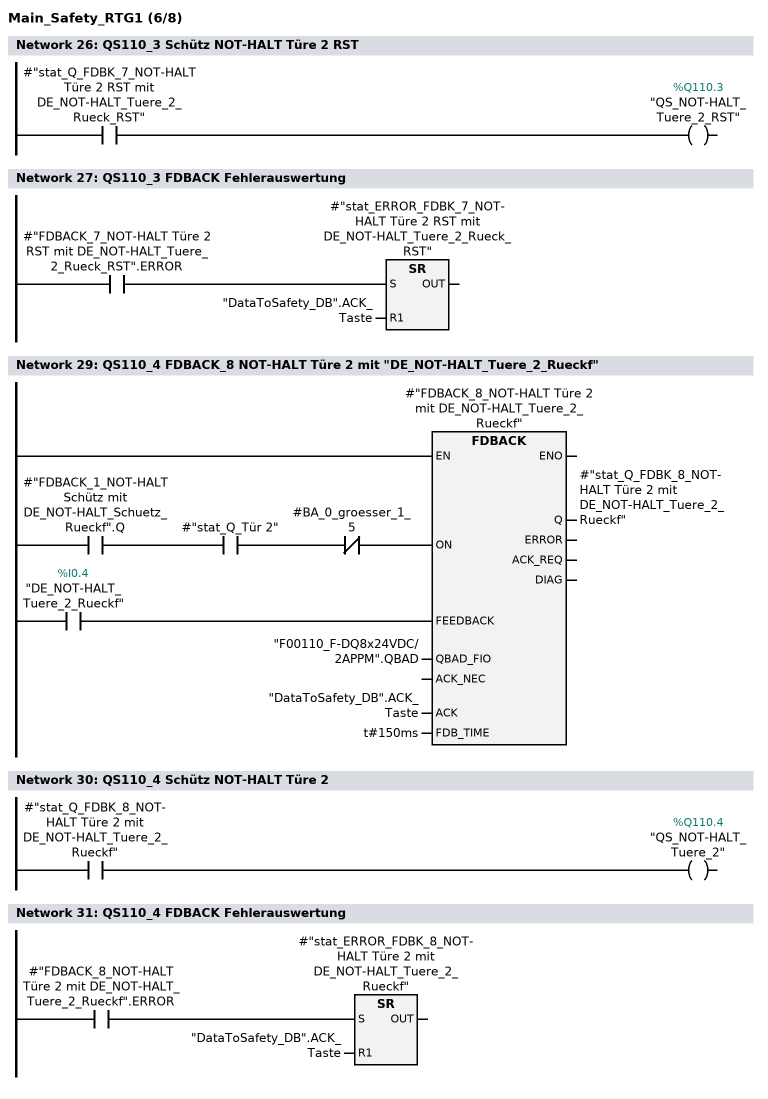
   RUNG wire#powerrail
      Contact( #"stat_Q_FDBK_7_NOT-HALT Türe 2 RST mit DE_NOT-HALT_Tuere_2_Rueck_RST" )
      Coil( "QS_NOT-HALT_Tuere_2_RST" )
   END_RUNG
   // the same network as SCL:
   "QS_NOT-HALT_Tuere_2_RST" := #"stat_Q_FDBK_7_NOT-HALT Türe 2 RST mit DE_NOT-HALT_Tuere_2_Rueck_RST";
END_REGION

REGION Network 27: QS110_3 FDBACK Fehlerauswertung
   RUNG wire#powerrail
      Contact( #"FDBACK_7_NOT-HALT Türe 2 RST mit DE_NOT-HALT_Tuere_2_Rueck_RST".ERROR )
      S_SR(operand := #"stat_ERROR_FDBK_7_NOT-HALT Türe 2 RST mit DE_NOT-HALT_Tuere_2_Rueck_RST", r1 := "DataToSafety_DB".ACK_Taste)
   END_RUNG
   // the same network as SCL:
   IF #"FDBACK_7_NOT-HALT Türe 2 RST mit DE_NOT-HALT_Tuere_2_Rueck_RST".ERROR THEN
       #"stat_ERROR_FDBK_7_NOT-HALT Türe 2 RST mit DE_NOT-HALT_Tuere_2_Rueck_RST" := TRUE;   // SR flip-flop
   END_IF;
   IF "DataToSafety_DB".ACK_Taste THEN
       #"stat_ERROR_FDBK_7_NOT-HALT Türe 2 RST mit DE_NOT-HALT_Tuere_2_Rueck_RST" := FALSE;
   END_IF;
END_REGION

REGION Network 28: *********************************************************************************************
END_REGION

REGION Network 29: QS110_4 FDBACK_8 NOT-HALT Türe 2 mit "DE_NOT-HALT_Tuere_2_Rueckf"
   RUNG wire#powerrail
      #"FDBACK_8_NOT-HALT Türe 2 mit DE_NOT-HALT_Tuere_2_Rueckf".FDBACK(ON := wire#w1, FEEDBACK := wire#w2, QBAD_FIO := "F00110_F-DQ8x24VDC/2APPM".QBAD, ACK_NEC :=, ACK := "DataToSafety_DB".ACK_Taste, FDB_TIME := t#150ms, Q => #"stat_Q_FDBK_8_NOT-HALT Türe 2 mit DE_NOT-HALT_Tuere_2_Rueckf", ERROR =>, ACK_REQ =>, DIAG =>)
   END_RUNG
   RUNG wire#powerrail
      Contact( #"FDBACK_1_NOT-HALT Schütz mit DE_NOT-HALT_Schuetz_Rueckf".Q )
      Contact( #"stat_Q_Tür 2" )
      I_Contact( #BA_0_groesser_1_5 )
   END_RUNG wire#w1
   RUNG wire#powerrail
      Contact( "DE_NOT-HALT_Tuere_2_Rueckf" )
   END_RUNG wire#w2
   // the same network as SCL:
   #"FDBACK_8_NOT-HALT Türe 2 mit DE_NOT-HALT_Tuere_2_Rueckf"(ON := #"FDBACK_1_NOT-HALT Schütz mit DE_NOT-HALT_Schuetz_Rueckf".Q AND #"stat_Q_Tür 2" AND NOT #BA_0_groesser_1_5,   // FDBACK
                           FEEDBACK := "DE_NOT-HALT_Tuere_2_Rueckf",
                           QBAD_FIO := "F00110_F-DQ8x24VDC/2APPM".QBAD,
                           ACK := "DataToSafety_DB".ACK_Taste,
                           FDB_TIME := t#150ms,
                           Q => #"stat_Q_FDBK_8_NOT-HALT Türe 2 mit DE_NOT-HALT_Tuere_2_Rueckf");
END_REGION

REGION Network 30: QS110_4 Schütz NOT-HALT Türe 2
   RUNG wire#powerrail
      Contact( #"stat_Q_FDBK_8_NOT-HALT Türe 2 mit DE_NOT-HALT_Tuere_2_Rueckf" )
      Coil( "QS_NOT-HALT_Tuere_2" )
   END_RUNG
   // the same network as SCL:
   "QS_NOT-HALT_Tuere_2" := #"stat_Q_FDBK_8_NOT-HALT Türe 2 mit DE_NOT-HALT_Tuere_2_Rueckf";
END_REGION

REGION Network 31: QS110_4 FDBACK Fehlerauswertung
   RUNG wire#powerrail
      Contact( #"FDBACK_8_NOT-HALT Türe 2 mit DE_NOT-HALT_Tuere_2_Rueckf".ERROR )
      S_SR(operand := #"stat_ERROR_FDBK_8_NOT-HALT Türe 2 mit DE_NOT-HALT_Tuere_2_Rueckf", r1 := "DataToSafety_DB".ACK_Taste)
   END_RUNG
   // the same network as SCL:
   IF #"FDBACK_8_NOT-HALT Türe 2 mit DE_NOT-HALT_Tuere_2_Rueckf".ERROR THEN
       #"stat_ERROR_FDBK_8_NOT-HALT Türe 2 mit DE_NOT-HALT_Tuere_2_Rueckf" := TRUE;   // SR flip-flop
   END_IF;
   IF "DataToSafety_DB".ACK_Taste THEN
       #"stat_ERROR_FDBK_8_NOT-HALT Türe 2 mit DE_NOT-HALT_Tuere_2_Rueckf" := FALSE;
   END_IF;
END_REGION

REGION Network 32: *********************************************************************************************
END_REGION

REGION Network 33: QS110_6 FDBACK_10 Sichere Bewegung
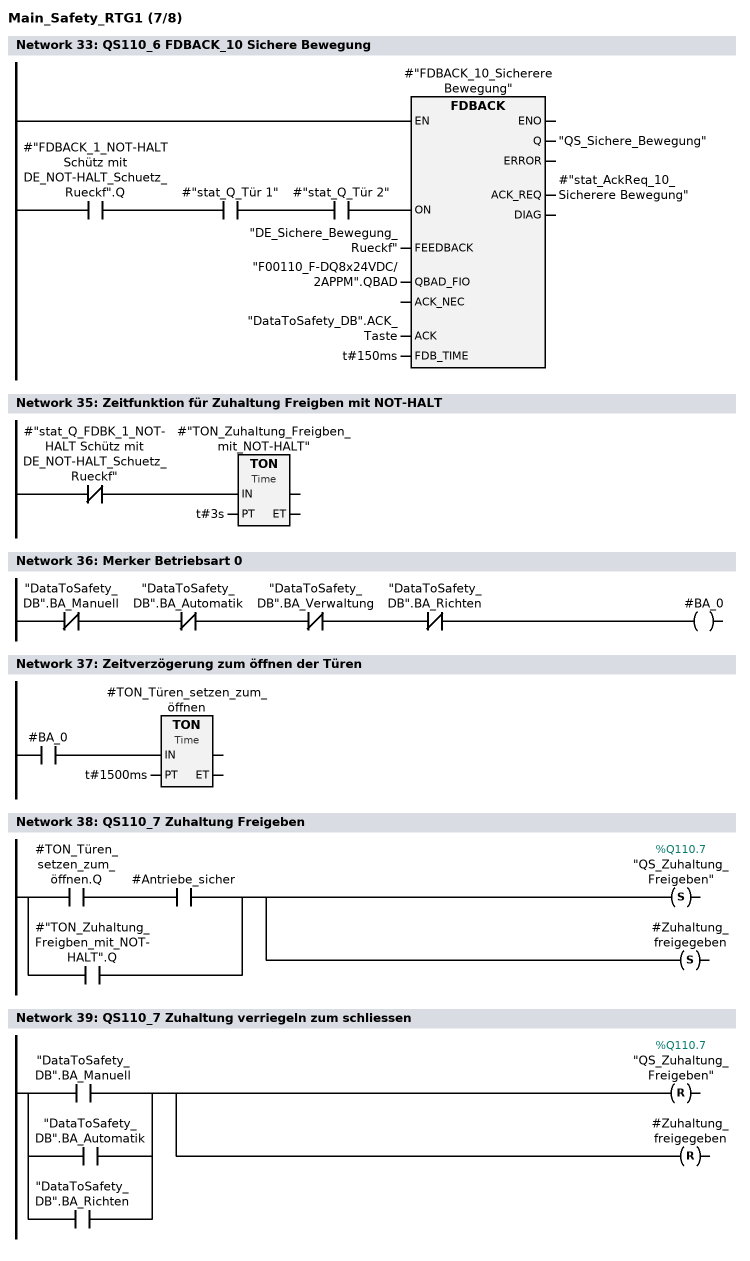
   RUNG wire#powerrail
      #"FDBACK_10_Sicherere Bewegung".FDBACK(ON := wire#w1, FEEDBACK := "DE_Sichere_Bewegung_Rueckf", QBAD_FIO := "F00110_F-DQ8x24VDC/2APPM".QBAD, ACK_NEC :=, ACK := "DataToSafety_DB".ACK_Taste, FDB_TIME := t#150ms, Q => "QS_Sichere_Bewegung", ERROR =>, ACK_REQ => #"stat_AckReq_10_Sicherere Bewegung", DIAG =>)
   END_RUNG
   RUNG wire#powerrail
      Contact( #"FDBACK_1_NOT-HALT Schütz mit DE_NOT-HALT_Schuetz_Rueckf".Q )
      Contact( #"stat_Q_Tür 1" )
      Contact( #"stat_Q_Tür 2" )
   END_RUNG wire#w1
   // the same network as SCL:
   #"FDBACK_10_Sicherere Bewegung"(ON := #"FDBACK_1_NOT-HALT Schütz mit DE_NOT-HALT_Schuetz_Rueckf".Q AND #"stat_Q_Tür 1" AND #"stat_Q_Tür 2",   // FDBACK
                           FEEDBACK := "DE_Sichere_Bewegung_Rueckf",
                           QBAD_FIO := "F00110_F-DQ8x24VDC/2APPM".QBAD,
                           ACK := "DataToSafety_DB".ACK_Taste,
                           FDB_TIME := t#150ms,
                           Q => "QS_Sichere_Bewegung",
                           ACK_REQ => #"stat_AckReq_10_Sicherere Bewegung");
END_REGION

REGION Network 34: *********************************************************************************************
END_REGION

REGION Network 35: Zeitfunktion für Zuhaltung Freigben mit NOT-HALT
   RUNG wire#powerrail
      I_Contact( #"stat_Q_FDBK_1_NOT-HALT Schütz mit DE_NOT-HALT_Schuetz_Rueckf" )
      { S7_Templates := "[time_type := Time, codedbool_type := DInt]" } #"TON_Zuhaltung_Freigben_mit_NOT-HALT".TON(pt := t#3s, et =>)
   END_RUNG
   // the same network as SCL:
   #"TON_Zuhaltung_Freigben_mit_NOT-HALT".TON(IN := NOT #"stat_Q_FDBK_1_NOT-HALT Schütz mit DE_NOT-HALT_Schuetz_Rueckf",
                           PT := t#3s);
END_REGION

REGION Network 36: Merker Betriebsart 0
   RUNG wire#powerrail
      I_Contact( "DataToSafety_DB".BA_Manuell )
      I_Contact( "DataToSafety_DB".BA_Automatik )
      I_Contact( "DataToSafety_DB".BA_Verwaltung )
      I_Contact( "DataToSafety_DB".BA_Richten )
      Coil( #BA_0 )
   END_RUNG
   // the same network as SCL:
   #BA_0 := NOT "DataToSafety_DB".BA_Manuell AND NOT "DataToSafety_DB".BA_Automatik AND NOT "DataToSafety_DB".BA_Verwaltung AND NOT "DataToSafety_DB".BA_Richten;
END_REGION

REGION Network 37: Zeitverzögerung zum öffnen der Türen
   RUNG wire#powerrail
      Contact( #BA_0 )
      { S7_Templates := "[time_type := Time, codedbool_type := DInt]" } #TON_Türen_setzen_zum_öffnen.TON(pt := t#1500ms, et =>)
   END_RUNG
   // the same network as SCL:
   #TON_Türen_setzen_zum_öffnen.TON(IN := #BA_0, PT := t#1500ms);
END_REGION

REGION Network 38: QS110_7 Zuhaltung Freigeben
   RUNG wire#powerrail
      Contact( #TON_Türen_setzen_zum_öffnen.Q )
      Contact( #Antriebe_sicher )
      wire#w1
      S_Coil( "QS_Zuhaltung_Freigeben" )
   END_RUNG
   RUNG wire#powerrail
      Contact( #"TON_Zuhaltung_Freigben_mit_NOT-HALT".Q )
   END_RUNG wire#w1
   RUNG wire#w1
      S_Coil( #Zuhaltung_freigegeben )
   END_RUNG
   // the same network as SCL:
   IF (#TON_Türen_setzen_zum_öffnen.Q AND #Antriebe_sicher) OR #"TON_Zuhaltung_Freigben_mit_NOT-HALT".Q THEN
       "QS_Zuhaltung_Freigeben" := TRUE;
       #Zuhaltung_freigegeben := TRUE;
   END_IF;
END_REGION

REGION Network 39: QS110_7 Zuhaltung verriegeln zum schliessen
   RUNG wire#powerrail
      Contact( "DataToSafety_DB".BA_Manuell )
      wire#w1
      R_Coil( "QS_Zuhaltung_Freigeben" )
   END_RUNG
   RUNG wire#powerrail
      Contact( "DataToSafety_DB".BA_Automatik )
   END_RUNG wire#w1
   RUNG wire#powerrail
      Contact( "DataToSafety_DB".BA_Richten )
   END_RUNG wire#w1
   RUNG wire#w1
      R_Coil( #Zuhaltung_freigegeben )
   END_RUNG
   // the same network as SCL:
   IF "DataToSafety_DB".BA_Manuell OR "DataToSafety_DB".BA_Automatik OR "DataToSafety_DB".BA_Richten THEN
       "QS_Zuhaltung_Freigeben" := FALSE;
       #Zuhaltung_freigegeben := FALSE;
   END_IF;
END_REGION

REGION Network 40: *********************************************************************************************
END_REGION

REGION Network 41: Global acknowledgment of all F-I/O in an F-runtime group
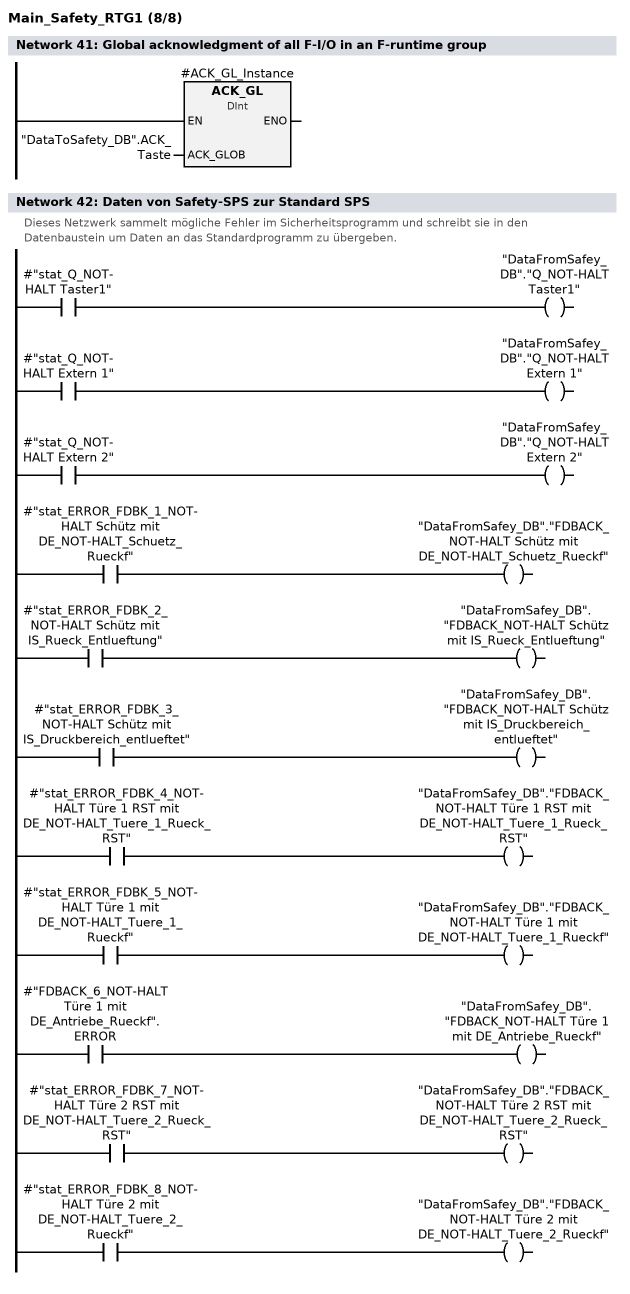
   RUNG wire#powerrail
      { S7_Templates := "codedbool_type := DInt" } #ACK_GL_Instance.ACK_GL(ACK_GLOB := "DataToSafety_DB".ACK_Taste)
   END_RUNG
   // the same network as SCL:
   #ACK_GL_Instance(ACK_GLOB := "DataToSafety_DB".ACK_Taste);   // ACK_GL
END_REGION

REGION Network 42: Daten von Safety-SPS zur Standard SPS
   // Dieses Netzwerk sammelt mögliche Fehler im Sicherheitsprogramm und schreibt sie in den Datenbaustein um Daten an das Standardprogramm zu übergeben.
   RUNG wire#powerrail
      Contact( #"stat_Q_NOT-HALT Taster1" )
      Coil( "DataFromSafey_DB"."Q_NOT-HALT Taster1" )
   END_RUNG
   RUNG wire#powerrail
      Contact( #"stat_Q_NOT-HALT Extern 1" )
      Coil( "DataFromSafey_DB"."Q_NOT-HALT Extern 1" )
   END_RUNG
   RUNG wire#powerrail
      Contact( #"stat_Q_NOT-HALT Extern 2" )
      Coil( "DataFromSafey_DB"."Q_NOT-HALT Extern 2" )
   END_RUNG
   RUNG wire#powerrail
      Contact( #"stat_ERROR_FDBK_1_NOT-HALT Schütz mit DE_NOT-HALT_Schuetz_Rueckf" )
      Coil( "DataFromSafey_DB"."FDBACK_NOT-HALT Schütz mit DE_NOT-HALT_Schuetz_Rueckf" )
   END_RUNG
   RUNG wire#powerrail
      Contact( #"stat_ERROR_FDBK_2_NOT-HALT Schütz mit IS_Rueck_Entlueftung" )
      Coil( "DataFromSafey_DB"."FDBACK_NOT-HALT Schütz mit IS_Rueck_Entlueftung" )
   END_RUNG
   RUNG wire#powerrail
      Contact( #"stat_ERROR_FDBK_3_NOT-HALT Schütz mit IS_Druckbereich_entlueftet" )
      Coil( "DataFromSafey_DB"."FDBACK_NOT-HALT Schütz mit IS_Druckbereich_entlueftet" )
   END_RUNG
   RUNG wire#powerrail
      Contact( #"stat_ERROR_FDBK_4_NOT-HALT Türe 1 RST mit DE_NOT-HALT_Tuere_1_Rueck_RST" )
      Coil( "DataFromSafey_DB"."FDBACK_NOT-HALT Türe 1 RST mit DE_NOT-HALT_Tuere_1_Rueck_RST" )
   END_RUNG
   RUNG wire#powerrail
      Contact( #"stat_ERROR_FDBK_5_NOT-HALT Türe 1 mit DE_NOT-HALT_Tuere_1_Rueckf" )
      Coil( "DataFromSafey_DB"."FDBACK_NOT-HALT Türe 1 mit DE_NOT-HALT_Tuere_1_Rueckf" )
   END_RUNG
   RUNG wire#powerrail
      Contact( #"FDBACK_6_NOT-HALT Türe 1 mit DE_Antriebe_Rueckf".ERROR )
      Coil( "DataFromSafey_DB"."FDBACK_NOT-HALT Türe 1 mit DE_Antriebe_Rueckf" )
   END_RUNG
   RUNG wire#powerrail
      Contact( #"stat_ERROR_FDBK_7_NOT-HALT Türe 2 RST mit DE_NOT-HALT_Tuere_2_Rueck_RST" )
      Coil( "DataFromSafey_DB"."FDBACK_NOT-HALT Türe 2 RST mit DE_NOT-HALT_Tuere_2_Rueck_RST" )
   END_RUNG
   RUNG wire#powerrail
      Contact( #"stat_ERROR_FDBK_8_NOT-HALT Türe 2 mit DE_NOT-HALT_Tuere_2_Rueckf" )
      Coil( "DataFromSafey_DB"."FDBACK_NOT-HALT Türe 2 mit DE_NOT-HALT_Tuere_2_Rueckf" )
   END_RUNG
   // the same network as SCL:
   "DataFromSafey_DB"."Q_NOT-HALT Taster1" := #"stat_Q_NOT-HALT Taster1";
   "DataFromSafey_DB"."Q_NOT-HALT Extern 1" := #"stat_Q_NOT-HALT Extern 1";
   "DataFromSafey_DB"."Q_NOT-HALT Extern 2" := #"stat_Q_NOT-HALT Extern 2";
   "DataFromSafey_DB"."FDBACK_NOT-HALT Schütz mit DE_NOT-HALT_Schuetz_Rueckf" := #"stat_ERROR_FDBK_1_NOT-HALT Schütz mit DE_NOT-HALT_Schuetz_Rueckf";
   "DataFromSafey_DB"."FDBACK_NOT-HALT Schütz mit IS_Rueck_Entlueftung" := #"stat_ERROR_FDBK_2_NOT-HALT Schütz mit IS_Rueck_Entlueftung";
   "DataFromSafey_DB"."FDBACK_NOT-HALT Schütz mit IS_Druckbereich_entlueftet" := #"stat_ERROR_FDBK_3_NOT-HALT Schütz mit IS_Druckbereich_entlueftet";
   "DataFromSafey_DB"."FDBACK_NOT-HALT Türe 1 RST mit DE_NOT-HALT_Tuere_1_Rueck_RST" := #"stat_ERROR_FDBK_4_NOT-HALT Türe 1 RST mit DE_NOT-HALT_Tuere_1_Rueck_RST";
   "DataFromSafey_DB"."FDBACK_NOT-HALT Türe 1 mit DE_NOT-HALT_Tuere_1_Rueckf" := #"stat_ERROR_FDBK_5_NOT-HALT Türe 1 mit DE_NOT-HALT_Tuere_1_Rueckf";
   "DataFromSafey_DB"."FDBACK_NOT-HALT Türe 1 mit DE_Antriebe_Rueckf" := #"FDBACK_6_NOT-HALT Türe 1 mit DE_Antriebe_Rueckf".ERROR;
   "DataFromSafey_DB"."FDBACK_NOT-HALT Türe 2 RST mit DE_NOT-HALT_Tuere_2_Rueck_RST" := #"stat_ERROR_FDBK_7_NOT-HALT Türe 2 RST mit DE_NOT-HALT_Tuere_2_Rueck_RST";
   "DataFromSafey_DB"."FDBACK_NOT-HALT Türe 2 mit DE_NOT-HALT_Tuere_2_Rueckf" := #"stat_ERROR_FDBK_8_NOT-HALT Türe 2 mit DE_NOT-HALT_Tuere_2_Rueckf";
END_REGION
END_FUNCTION_BLOCK

FUNCTION_BLOCK "08_Systemzeit"   // FB167, LAD
{ S7_Optimized_Access := 'TRUE' }
// stored: MemoryReserve 100, SetENOAutomatically false
   VAR
      outputTIME : Date_And_Time;
      returnValue : Int;
      inputTIME : Date_And_Time;
      returnValueT : Int;
      execute : Bool;
   END_VAR
BEGIN

REGION Network 1: Aktuelles Datum und Uhrzeit auslesen
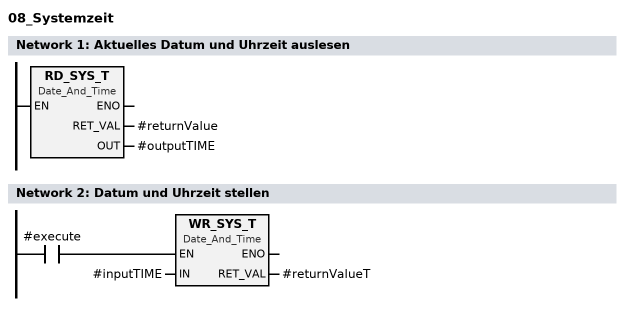
   RUNG wire#powerrail
      { S7_Templates := "date_type := Date_And_Time" } RD_SYS_T(RET_VAL => #returnValue, OUT => #outputTIME)
   END_RUNG
   // the same network as SCL:
   #returnValue := RD_SYS_T(OUT => #outputTIME);
END_REGION

REGION Network 2: Datum und Uhrzeit stellen
   RUNG wire#powerrail
      Contact( #execute )
      { S7_Templates := "date_type := Date_And_Time" } WR_SYS_T(IN := #inputTIME, RET_VAL => #returnValueT)
   END_RUNG
   // the same network as SCL:
   IF #execute THEN #returnValueT := WR_SYS_T(IN := #inputTIME); END_IF;
END_REGION
END_FUNCTION_BLOCK

FUNCTION "AchsePOS_BIT" : Void   // FC109, STL
TITLE = Achsenposition IST-POS mit Vorgabe vergleichen und Bit setzen
{ S7_Optimized_Access := 'FALSE' }
// stored: AutoNumber false
   VAR_INPUT
      ISTPOS_Achse : Real;   // Istposition der Achse
      POS_Vorgabe : Real;   // Achsposition die als Bit-Position benötigt wird
      Max_Abweichung : Real;   // +/- Abweichung in mm zur Achsposition
   END_VAR
   VAR_OUTPUT
      POS_OK : Bool;   // Wenn Istposition im Fenster POS_Vorgabe +/- MAX Abweichung ist dann VKE=1
   END_VAR
BEGIN

NETWORK
TITLE = Wenn Istposition im Fenster POS_Vorgabe +/- MAX Abweichung ist dann VKE=1
      A(;
      L     #ISTPOS_Achse;
      L     #POS_Vorgabe;
      -R;
      ABS;
      L     #Max_Abweichung;
      <=R;
      );
      =     #POS_OK;
END_FUNCTION

FUNCTION_BLOCK "Drehtelleransteuerung"   // FB117, STL
TITLE = Drehteller Ansteuerung über Schütz, Abfrage Endschalter
{ S7_Optimized_Access := 'TRUE' }
// stored: AutoNumber false, MemoryReserve 100
   VAR_INPUT
      ES_GS : Bool;
      ES_Motor_aus : Bool;
      Automatik : Bool;
      Manuell : Bool;
      Einrichten : Bool;
      Ablauf_aktiv : Bool;
      Richten : Bool;
      SM_reset : Bool;
      Reset_Frg : Bool;
      Not_Aus_OK : Bool;
      Tueren_OK : Bool;
      Lichtvorhang_OK : Bool;
      Sicherheitsbit_DT : Bool;
      TP_Taste_tippen : Bool;
      Start_taste_tippen : Bool;
      links0_rechts1_drehen : Bool;
      Richten_erforderlich : Bool;
      LVZ_Timer : Timer;
      Timer_ueberdrehen : Timer;
      SVZ : Timer;
   END_VAR
   VAR_OUTPUT
      Schuetz_links : Bool;
      Schuetz_rechts : Bool;
      DT_Bremse : Bool;
   END_VAR
   VAR_IN_OUT
      Freigabe_DT : Bool;
      Manuellfreigabe : Bool;
      Richtenfreigabe : Bool;
      Fertigmeldung_Drehteller : Bool;
      Betriebsfertigmeldung : Bool;
      SM_GS : Bool;
      SM_AS : Bool;
      SM_Wartung : Bool;
      Auto_Frg_GS : Bool;
      Auto_Frg_AS : Bool;
      Manu_Frg_GS : Bool;
      Manu_Frg_AS : Bool;
      Einr_Frg_GS : Bool;
      Einr_Frg_AS : Bool;
      Init_Frg_GS : Bool;
      Init_Frg_AS : Bool;
      Richt_Frg_GS : Bool;
      Richt_Frg_AS : Bool;
   END_VAR
   VAR
      SchrittA1 : Bool;
      SchrittA2 : Bool;
      SchrittA3 : Bool;
      HM_DT_Frg_loeschen : Bool;
      FP_DT_frg_loeschen : Bool;
      SchrittM1 : Bool;
      SchrittM2 : Bool;
      LV_unterbrochen : Bool;
      HM_Tippen : Bool;
      FP_Tippen : Bool;
      FP_Start_Tippen : Bool;
   END_VAR
BEGIN

NETWORK
TITLE = Störmeldungen
      A     #ES_GS;
      A     #SchrittA1;
      AN    #SchrittA2;
      O(;
      AN    #ES_GS;
      A     #SchrittA2;
      AN    #SchrittA3;
      );
      AN    #SM_reset;
      L     S5T#1S;
      SD    #LVZ_Timer;

      A     #LVZ_Timer;
      S     #SM_GS;


      AN    #ES_Motor_aus;
      A     #SchrittA1;
      AN    #SchrittA2;
      O(;
      A     #ES_Motor_aus;
      A     #SchrittA2;
      AN    #SchrittA3;
      );
      O(;
      AN    #ES_GS;
      A     #ES_Motor_aus;
      );
      AN    #SM_reset;
      L     S5T#1S;
      SD    #Timer_ueberdrehen;

      A     #Timer_ueberdrehen;
      S     #SM_AS;

      A     #SM_GS;
      A     #SM_reset;
      R     #SM_GS;

      A     #SM_AS;
      A     #SM_reset;
      R     #SM_AS;



NETWORK
TITLE = Lichtvorhang unterbrochen speichern
      A     #SchrittA1;
      AN    #Lichtvorhang_OK;
      S     #LV_unterbrochen;
      R     #SchrittA1;
      R     #SchrittA1;
      R     #SchrittA3;
      R     #DT_Bremse;
      R     #Schuetz_rechts;
      R     #Schuetz_links;



NETWORK
TITLE = Fertigmeldung DT
      A     #Betriebsfertigmeldung;
      FP    #HM_DT_Frg_loeschen;
      =     #FP_DT_frg_loeschen;

      A     #FP_DT_frg_loeschen;
      S     #Fertigmeldung_Drehteller;
      R     #Betriebsfertigmeldung;



NETWORK
TITLE = Sicherheitsabfragen
      A     #Not_Aus_OK;
      A     #Tueren_OK;
      A     #Lichtvorhang_OK;
      A     #Sicherheitsbit_DT;
      JCN   Ende;
      A     #Automatik;
      A     #Ablauf_aktiv;
      O;
      A     #Manuell;
      A     #Manuellfreigabe;
      O     #Richten_erforderlich;
      JC    M010;
      A     #Manuell;
      AN    #Manuellfreigabe;
      JC    M050;

      JU    Ende;



NETWORK
TITLE = Schritt1: Ansteuerung DT Automatik/Manuell
M010: A     #SchrittA1;
      JC    M020;
      A     #Freigabe_DT;
      A     #ES_GS;
//   UN    #ES_Motor_aus
      O     #Manuellfreigabe;
      O(;
      A     #Richten_erforderlich;
      A     #Richtenfreigabe;
      );
      O(;
      A     #Lichtvorhang_OK;
      A     #LV_unterbrochen;
      );
      AN    #SM_GS;
      AN    #SM_AS;
      S     #DT_Bremse;
      R     #Freigabe_DT;
      R     #Richtenfreigabe;
      R     #LV_unterbrochen;

      A     #DT_Bremse;
      A     #links0_rechts1_drehen;
      S     #Schuetz_rechts;

      A     #DT_Bremse;
      AN    #links0_rechts1_drehen;
      S     #Schuetz_links;

      A     #Schuetz_rechts;
      O     #Schuetz_links;
      A     #DT_Bremse;
      S     #SchrittA1;
      JC    M021;
      BEU;
M021: CLR;
      SD    #SVZ;
      BEU;



NETWORK
TITLE = Schritt2: ES_GS geht weg
M020: A     #SchrittA2;
      JC    M030;
      AN    #ES_GS;
      A     #ES_Motor_aus;
      O     #SM_GS;
      O     #SM_AS;
      S     #SchrittA2;
      JC    M031;
      BEU;
M031: CLR;
      SD    #SVZ;
      BEU;



NETWORK
TITLE = Schritt3: ES_GS kommt und ES_Motor_aus geht weg
M030: A     #SchrittA3;
      JC    M040;
      A     #ES_GS;
      A     #ES_Motor_aus;
      AN    #Richten_erforderlich;
      O(;
      A     #ES_Motor_aus;
      A     #ES_GS;
      A     #Richten_erforderlich;
      );
      O     #SM_GS;
      O     #SM_AS;
      O(;
      AN    #SM_GS;
      AN    #SM_AS;
      A     #ES_GS;
      AN    #ES_Motor_aus;
      A     #SM_reset;
      );
      R     #Schuetz_rechts;
      R     #Schuetz_links;
      R     #DT_Bremse;
      S     #Betriebsfertigmeldung;
      S     #SchrittA3;
      JC    M041;
      BEU;
M041: CLR;
      SD    #SVZ;
      BEU;



NETWORK
TITLE = Schrittkettenende
M040: SET;
      R     #SchrittA1;
      R     #SchrittA2;
      R     #SchrittA3;
      R     #Manuellfreigabe;
      BEU;



NETWORK
TITLE = Schritt1: Ansteuerung DT Manuell-Tippen
M050: A     #TP_Taste_tippen;
      A     #Start_taste_tippen;
      FP    #FP_Start_Tippen;
      S     #HM_Tippen;

      A(;
      A     #ES_GS;
      A     #ES_Motor_aus;
      FP    #FP_Tippen;
      );
      ON    #TP_Taste_tippen;
      ON    #Start_taste_tippen;
      R     #HM_Tippen;

      A     #HM_Tippen;
      =     #DT_Bremse;

      A     #DT_Bremse;
      A     #links0_rechts1_drehen;
      =     #Schuetz_rechts;

      A     #DT_Bremse;
      AN    #links0_rechts1_drehen;
      =     #Schuetz_links;

      BEU;



NETWORK
TITLE = Ende wenn nichts angewählt
Ende: NOP   0;
      SET;
      R     #DT_Bremse;
      R     #Schuetz_rechts;
      R     #Schuetz_links;
      R     #SchrittA1;
      R     #SchrittA2;
      R     #SchrittA3;
      R     #Manuellfreigabe;

      BEU;

END_FUNCTION_BLOCK

FUNCTION "Real Laden" : Void   // FC131, STL
TITLE = Real Laden für Graph
{ S7_Optimized_Access := 'FALSE' }
// stored: AutoNumber false
   VAR_INPUT
      Eingabewert : Real;
   END_VAR
   VAR_OUTPUT
      Ausgabewert : Real;
   END_VAR
BEGIN

NETWORK
TITLE = 
      L     #Eingabewert;
      T     #Ausgabewert;
END_FUNCTION

FUNCTION "Zählerfunktion mit STOP" : Void   // FC106, STL
TITLE = Zählerfunktion mit Stop
{ S7_Optimized_Access := 'FALSE' }
AUTHOR : SD
FAMILY : Zähler
// stored: AutoNumber false
   VAR_INPUT
      Stopwert : DInt;   // Bei diesem Wert wird ein Stopsignal ausgegeben
      RESET : Bool;
   END_VAR
   VAR_IN_OUT
      Zaehlsignal : Bool;
      Zaehlerstand : DInt;
      Stopbit : Bool;   // Stopbit
   END_VAR
BEGIN

NETWORK
TITLE = Zählsignal
      AN    #Zaehlsignal;
      JC    M031;

      SET;
      R     #Zaehlsignal;

NETWORK
TITLE = Zählerstand erhöhen
      L     #Zaehlerstand;
      L     1;
      +D;
      T     #Zaehlerstand;

NETWORK
TITLE = Vergleich von Ist und Sollstand
      L     #Zaehlerstand;
      L     #Stopwert;
      <D;
      JC    M031;
      SET;
      S     #Stopbit;

M031: NOP   0;

NETWORK
TITLE = Reset Stopbit und Zählerstand
      AN    #RESET;
      JC    M041;
      L     0;
      T     #Zaehlerstand;

      SET;
      R     #Stopbit;
M041: NOP   0;
END_FUNCTION

FUNCTION "GIT_Testbaustein in KOP" : Void   // FC5, LAD
{ S7_Optimized_Access := 'TRUE' }
// stored: SetENOAutomatically false
BEGIN

REGION Network 1
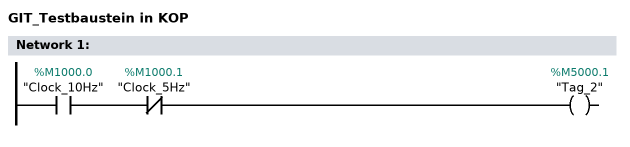
   RUNG wire#powerrail
      Contact( "Clock_10Hz" )
      I_Contact( "Clock_5Hz" )
      Coil( "Tag_2" )
   END_RUNG
   // the same network as SCL:
   "Tag_2" := "Clock_10Hz" AND NOT "Clock_5Hz";
END_REGION
END_FUNCTION

ORGANIZATION_BLOCK "IO access error"
{ S7_Optimized_Access := 'TRUE' }
VERSION : 0.1

BEGIN
END_ORGANIZATION_BLOCK

ORGANIZATION_BLOCK "Programming error"
{ S7_Optimized_Access := 'TRUE' }
VERSION : 0.1

BEGIN
END_ORGANIZATION_BLOCK

ORGANIZATION_BLOCK "Rack or station failure"
{ S7_Optimized_Access := 'TRUE' }
VERSION : 0.1

BEGIN
END_ORGANIZATION_BLOCK

ORGANIZATION_BLOCK "Startup"
TITLE = "Complete Restart"
{ S7_Optimized_Access := 'TRUE' }
VERSION : 0.1

BEGIN
END_ORGANIZATION_BLOCK

FUNCTION_BLOCK "BB_Ansteuerung_Afag_Dreh_V03.16"
TITLE = 'FB Positionierbetrieb'
{ S7_Optimized_Access := 'TRUE' }
AUTHOR : Essmann
FAMILY : metronix
NAME : position
VERSION : 1.1
//Der Baustein kann nicht rückübersetzt und unter STEP7 bearbeitet werden.  Der Baustein kann nur als Quelle im Ordner "Quellen" bearbeitet werden.    IO-Variablen  
   VAR_INPUT 
      E_UDT_Afag_ist_Werte : "Afag_ist_Werte";
      E_BA_Manuell : Bool;
      E_I_Manuell_Geschwindigkeit_Prozent : Int;
      E_Richten_reset_FRG : Bool;
      E_drive_enable : Bool := FALSE;
      E_start_homing : Bool := FALSE;
      E_change_immediatly : Bool := FALSE;
      E_intermediate_stop : Bool := FALSE;
      E_hold : Bool := FALSE;
      E_jog_pos : Bool := FALSE;
      E_jog_neg : Bool := FALSE;
      E_fault_reset : Bool := FALSE;
      E_Tipp_pos : Bool;
      E_Tipp_neg : Bool;
      E_Start_pos_man : Bool;
      E_R_Verfahrweg_Grad : Real;
      E_R_Afag_soll_wert_man_Grad : Real;
      E_I_Max_Speed_Grad_s : Int;
      E_I_Max_Beschleunigung_Grad_s : Int;
   END_VAR

   VAR_OUTPUT 
      A_drive_enable_ok : Bool := FALSE;
      A_home_valid : Bool := FALSE;
      A_pos_ok : Bool := FALSE;
      A_velo_zero : Bool := FALSE;
      A_fault : Bool := FALSE;   // statische Variablen
      A_Fahrauftrag_Aktiv : Bool;
      A_Afag_ist_wert_Grad : Real;
   END_VAR

   VAR_IN_OUT 
      E_A_UDT_Afag_Positionen : "Afag_Variablen_Positionen_Dreh";
      A_UDT_Afag_soll_Werte : "Afag_soll_Werte";
   END_VAR

